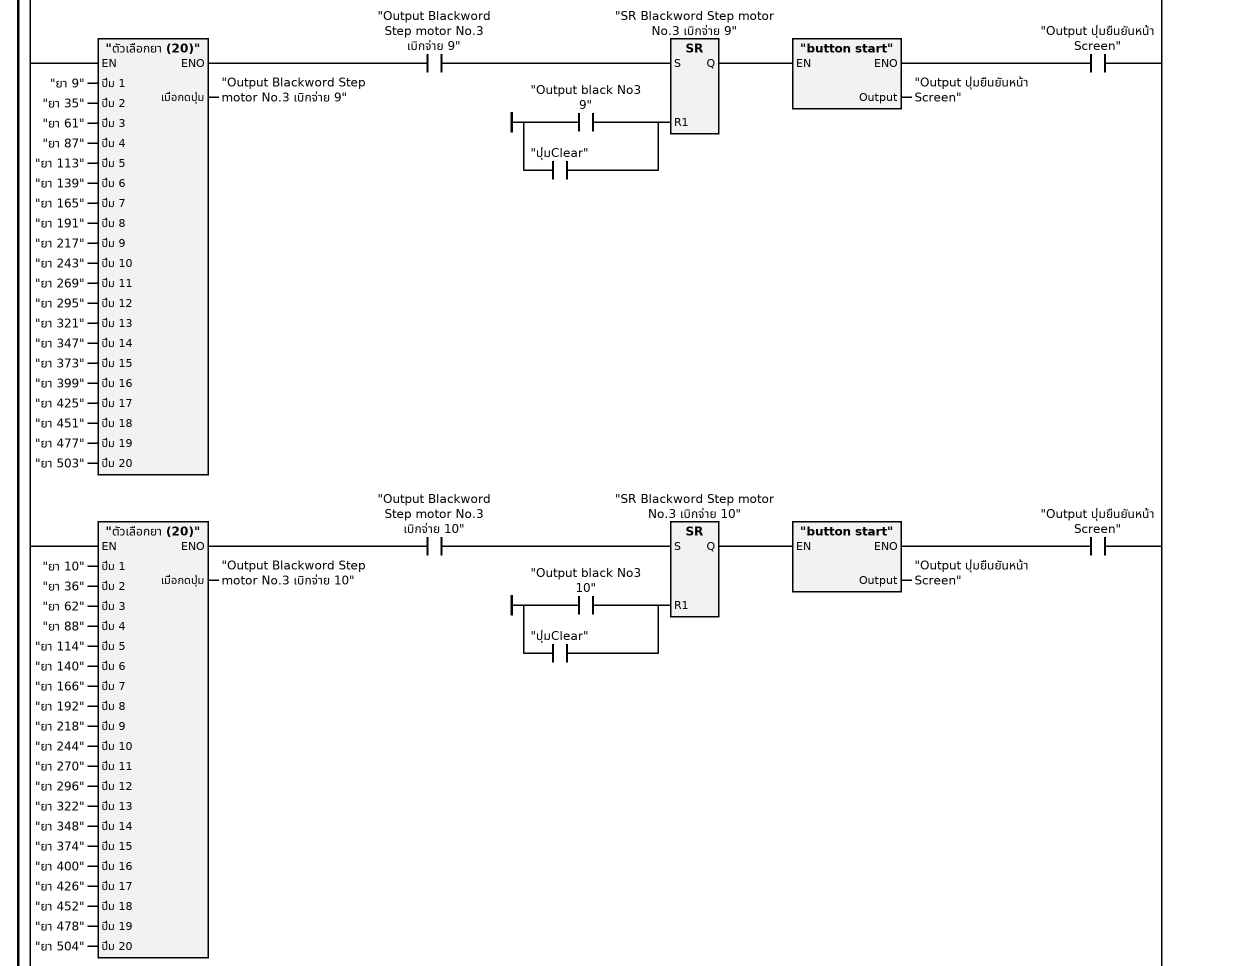
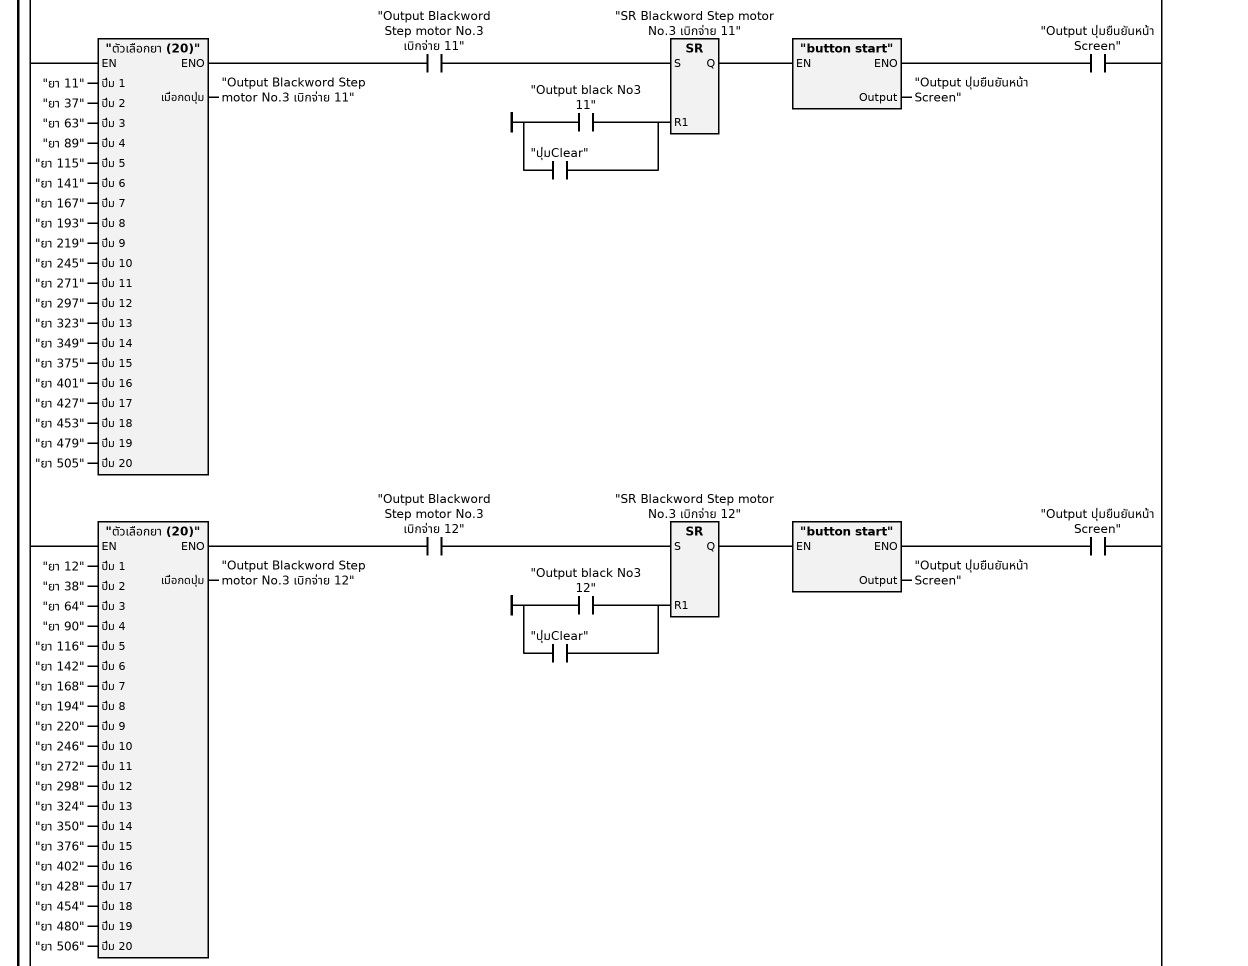
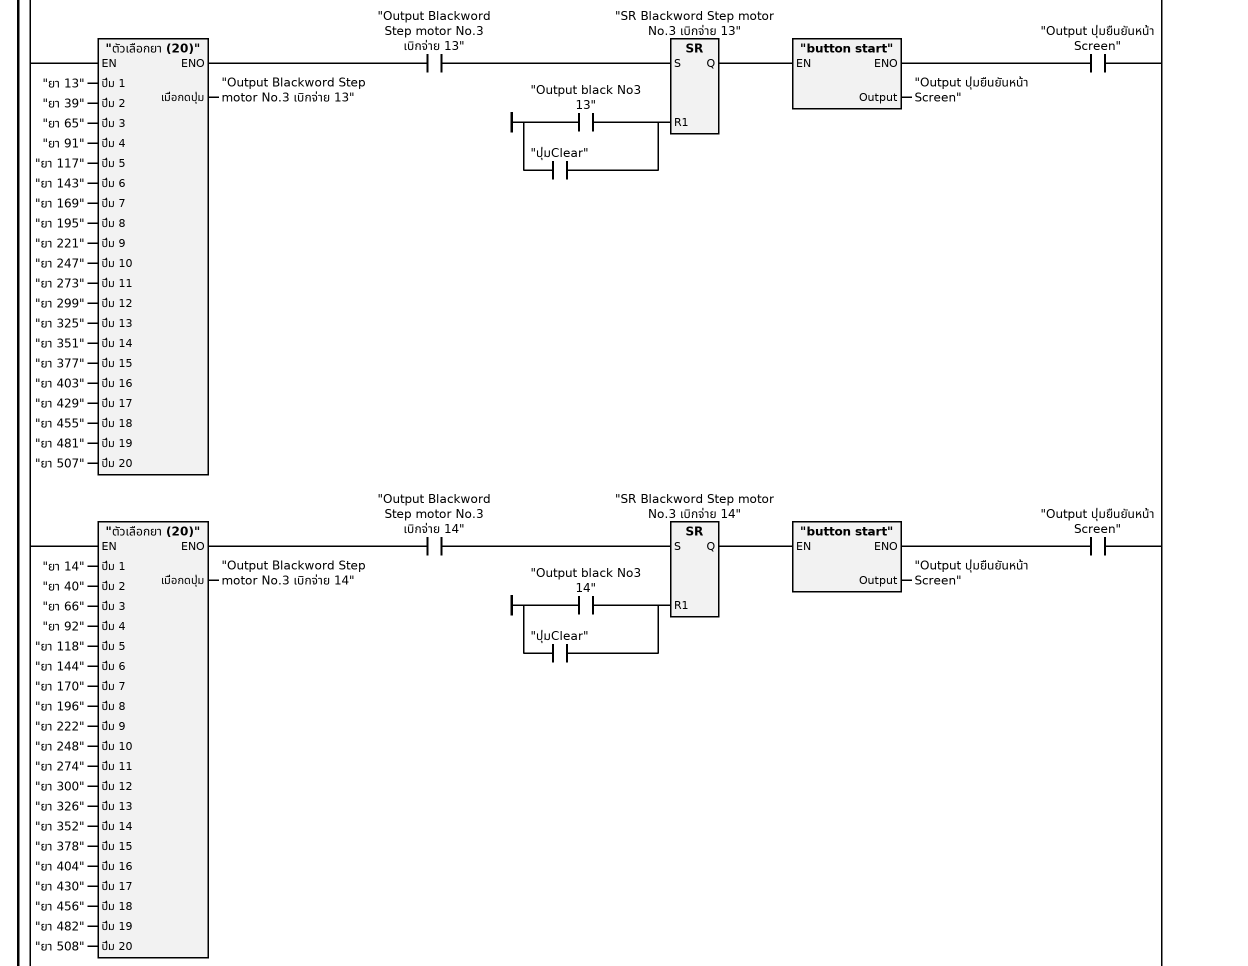
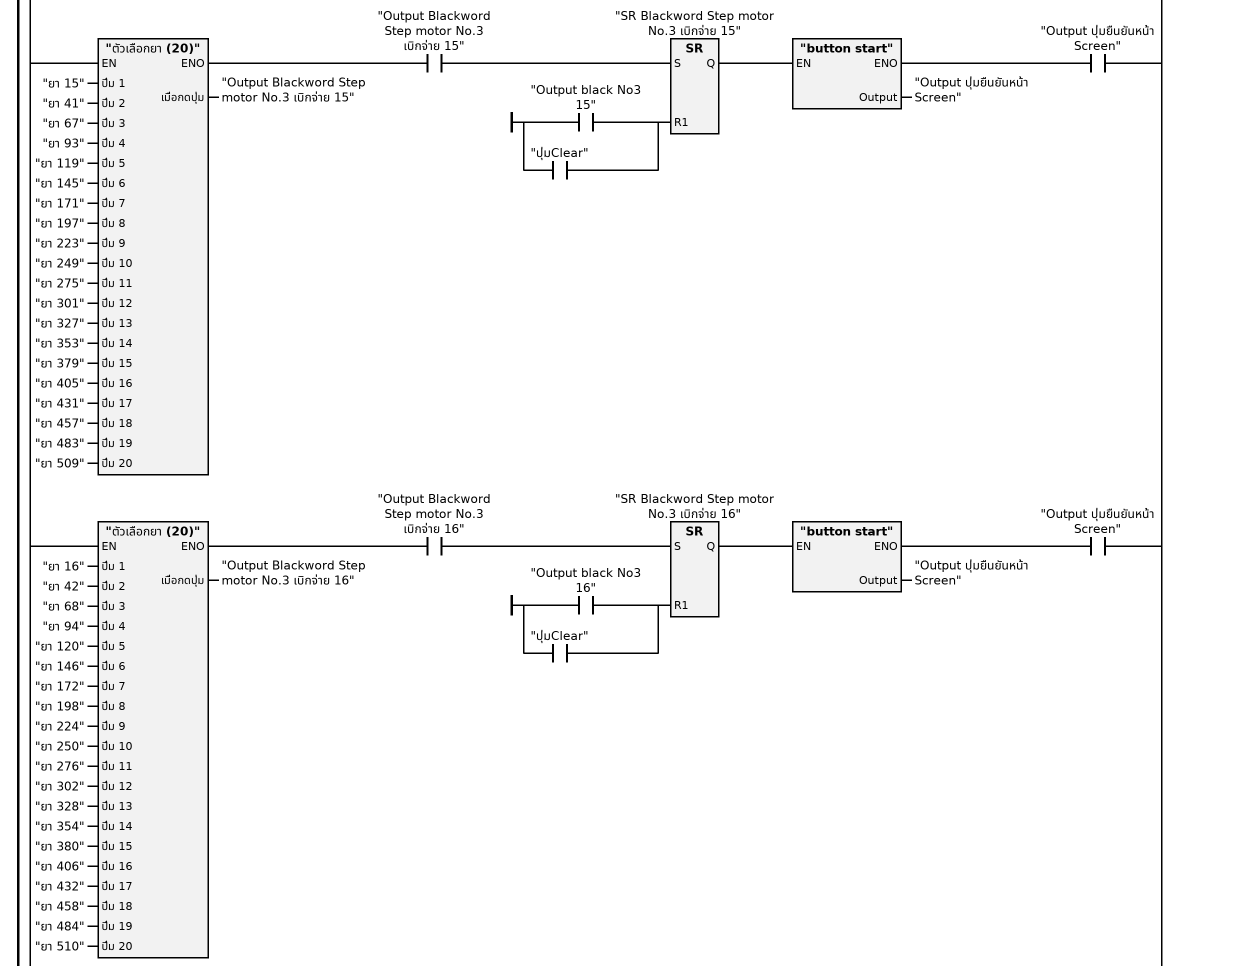
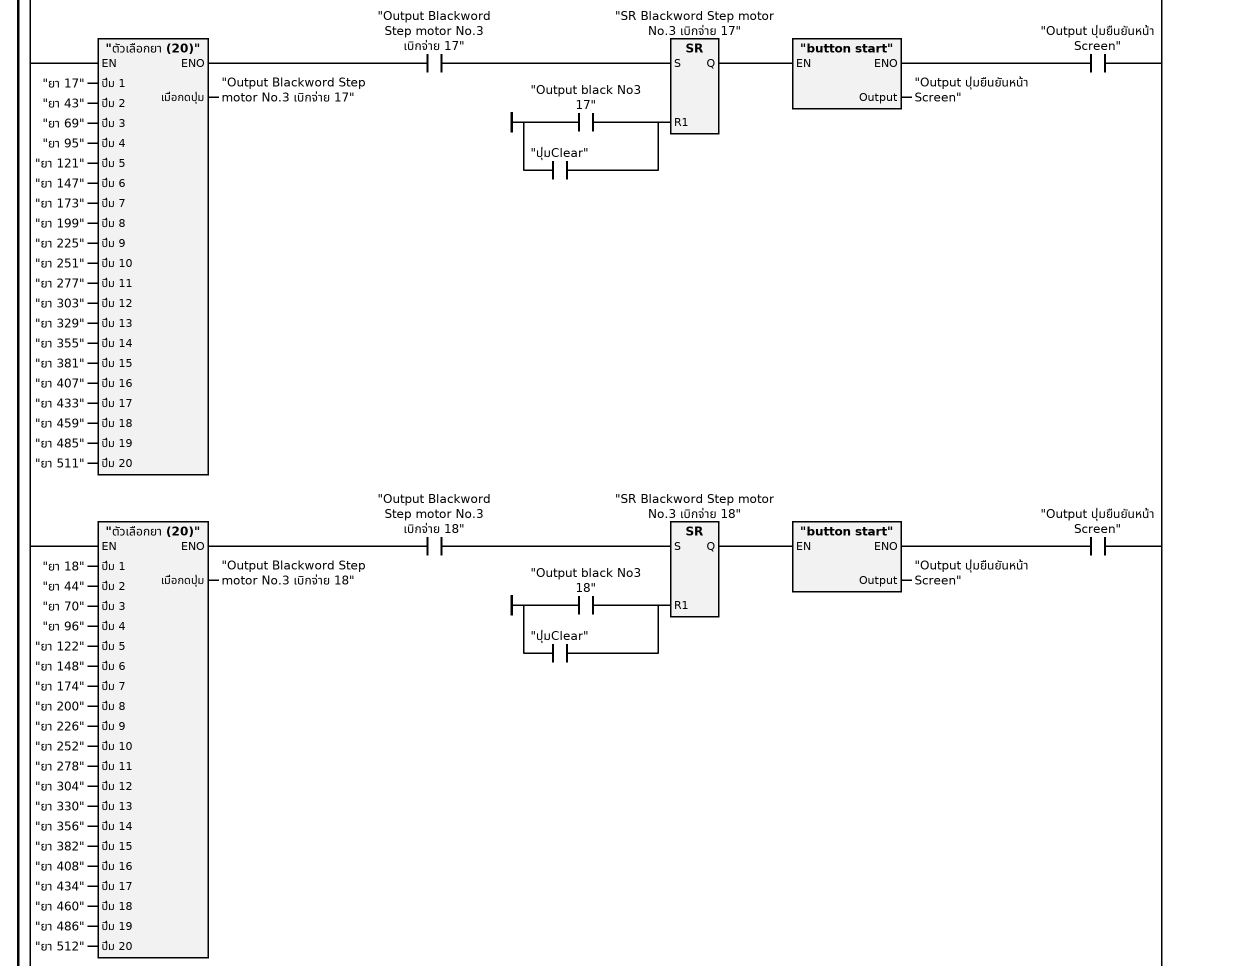
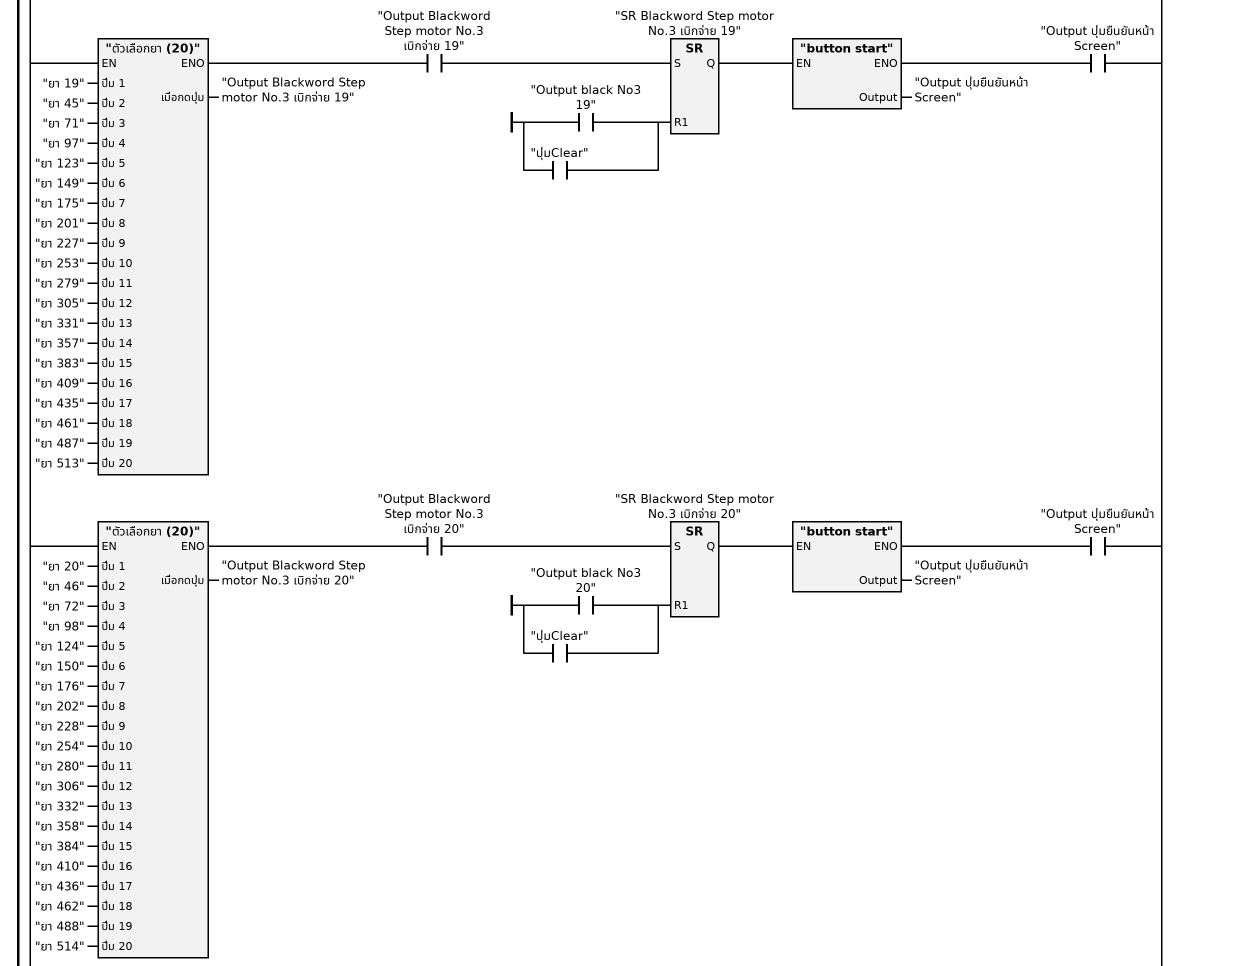
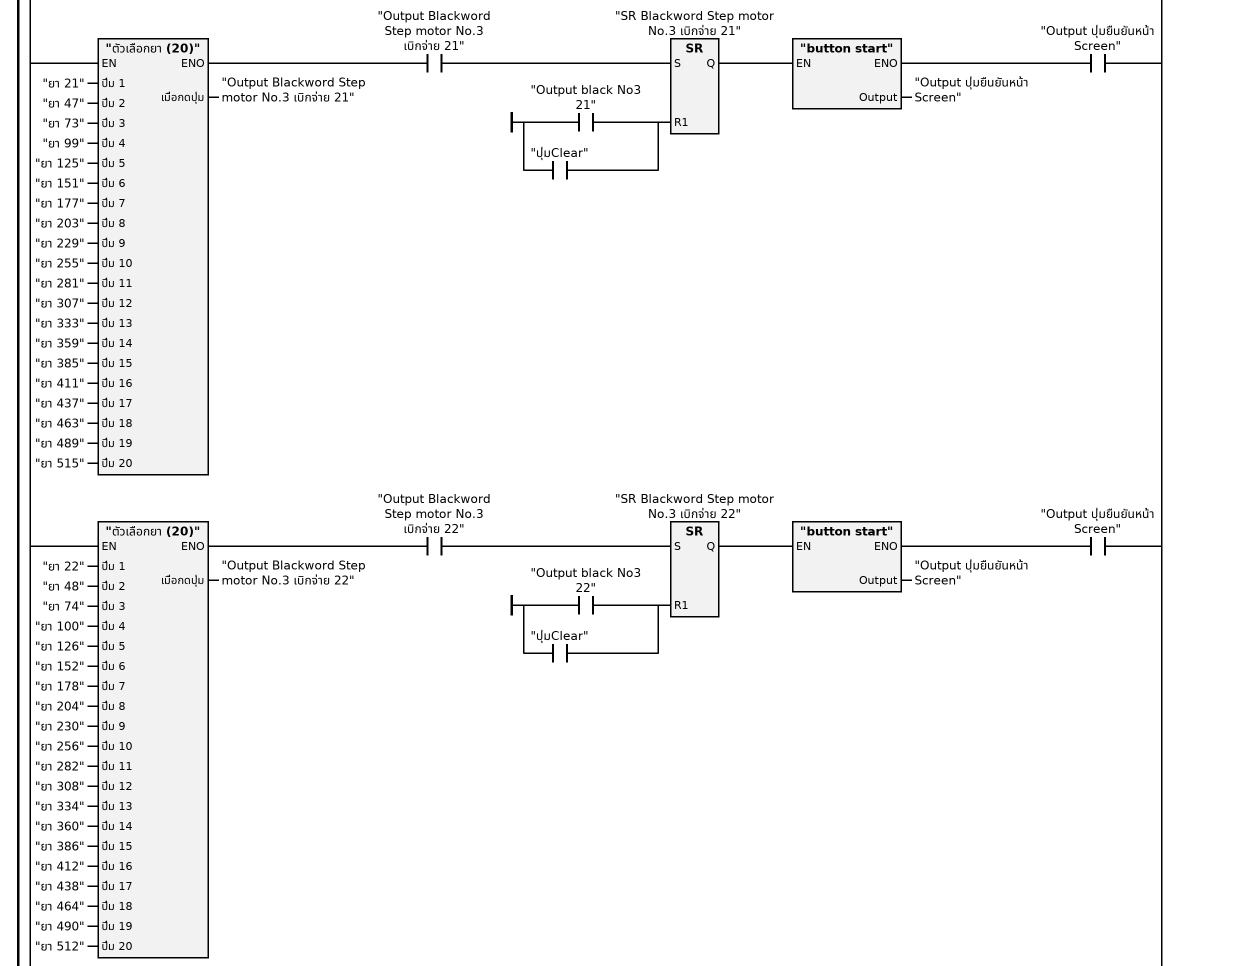
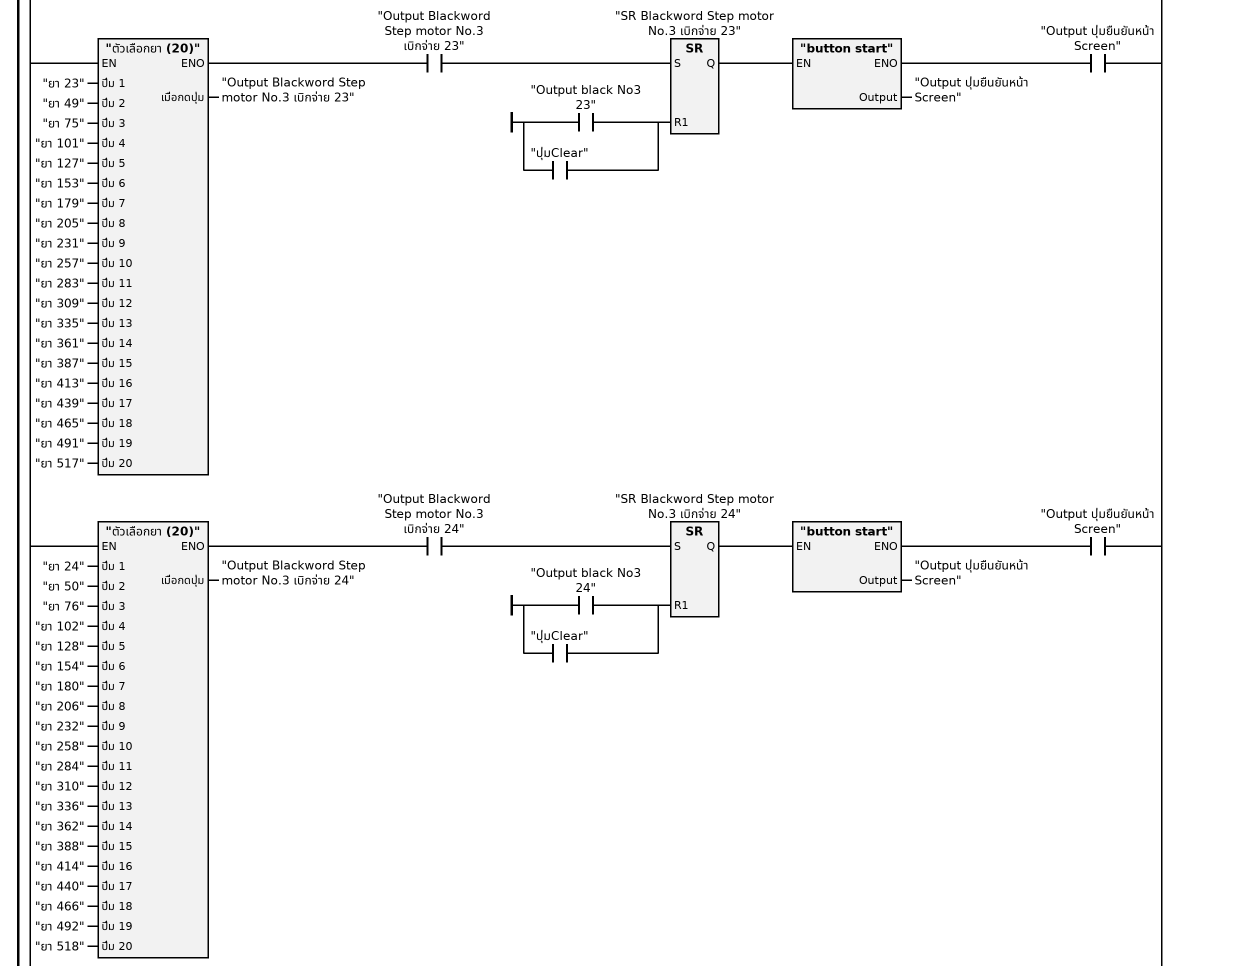
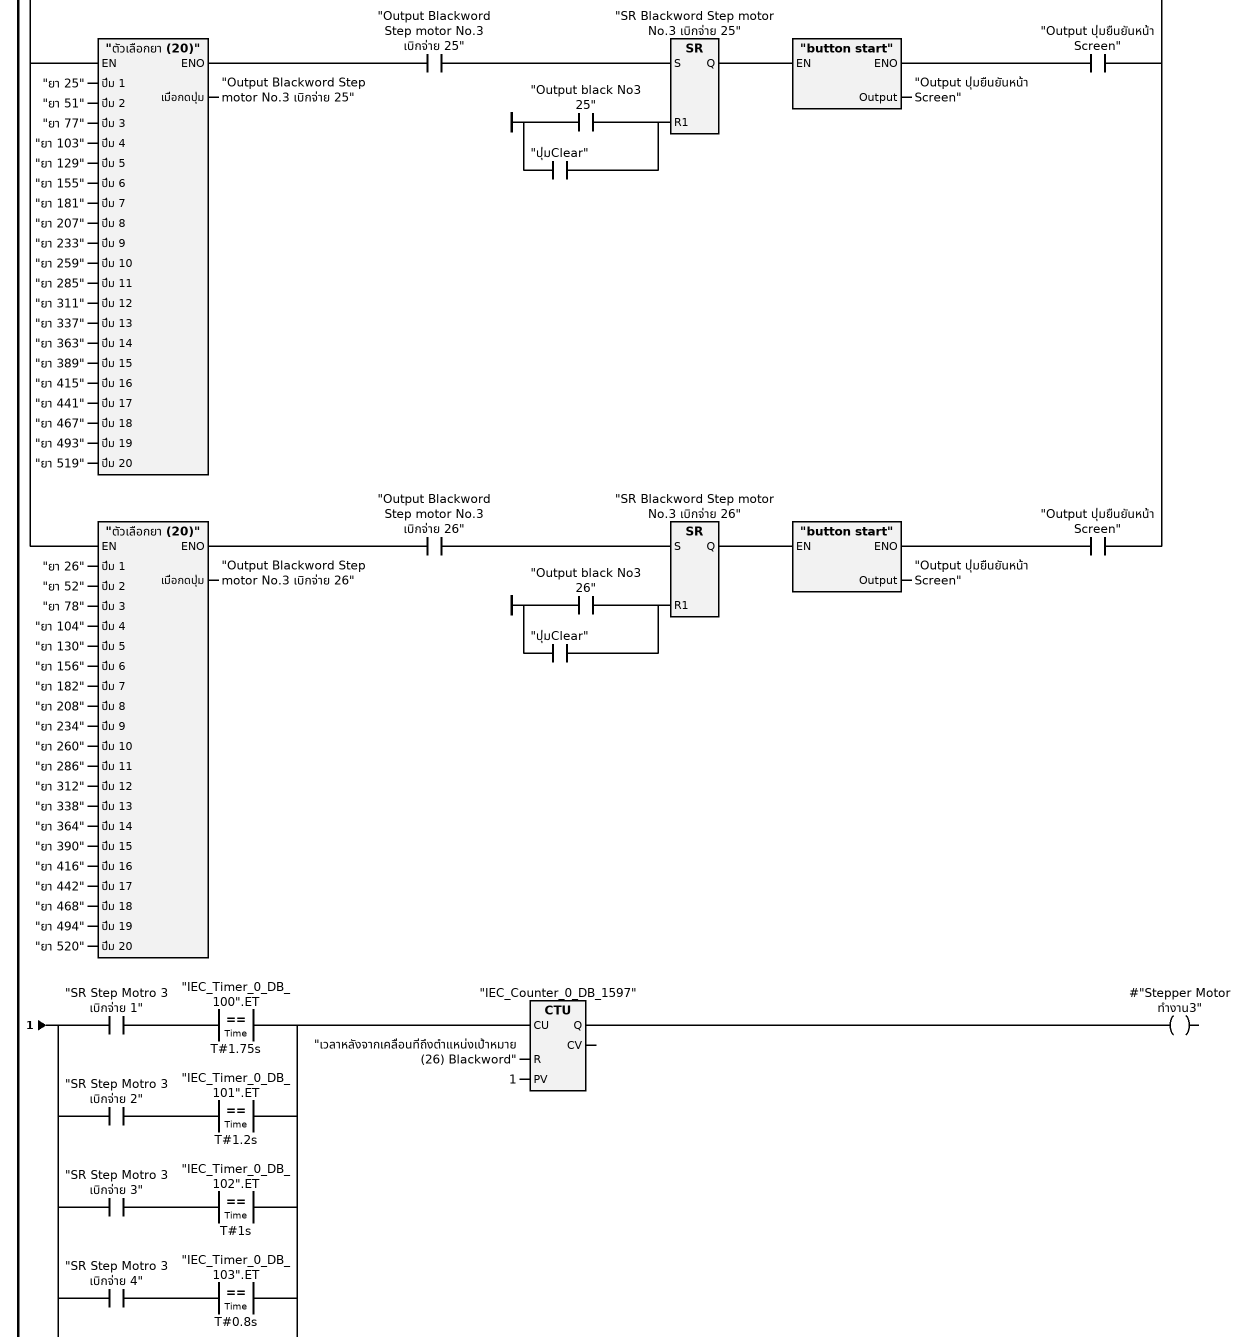
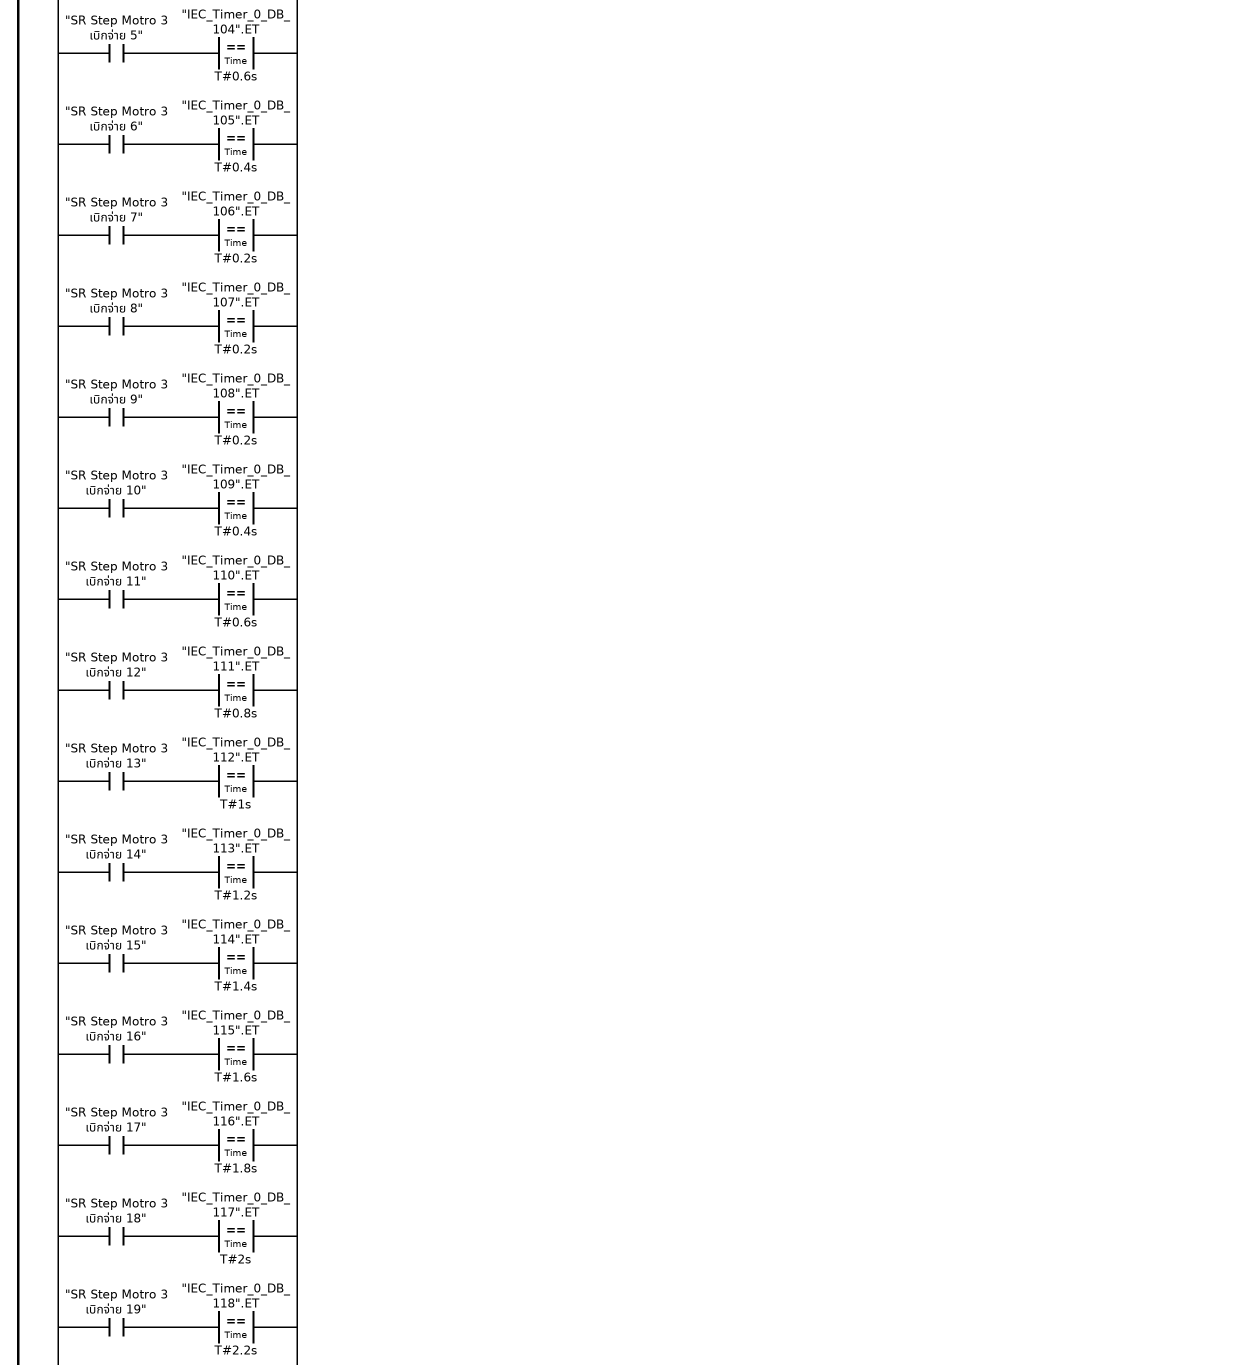
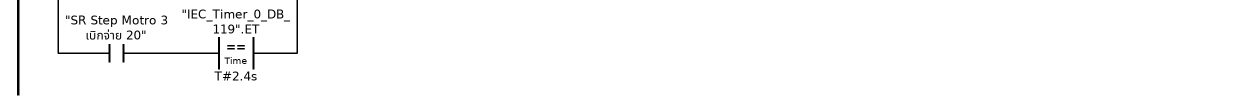
   "ตัวเลือกยา (20)"("ปึ่ม 1" := "ยา 1",
                     "ปึ่ม 2" := "ยา 27",
                     "ปึ่ม 3" := "ยา 53",
                     "ปึ่ม 4" := "ยา 79",
                     "ปึ่ม 5" := "ยา 105",
                     "ปึ่ม 6" := "ยา 131",
                     "ปึ่ม 7" := "ยา 157",
                     "ปึ่ม 8" := "ยา 183",
                     "ปึ่ม 9" := "ยา 209",
                     "ปึ่ม 10" := "ยา 235",
                     "ปึ่ม 11" := "ยา 261",
                     "ปึ่ม 12" := "ยา 287",
                     "ปึ่ม 13" := "ยา 313",
                     "ปึ่ม 14" := "ยา 339",
                     "ปึ่ม 15" := "ยา 365",
                     "ปึ่ม 16" := "ยา 391",
                     "ปึ่ม 17" := "ยา 417",
                     "ปึ่ม 18" := "ยา 443",
                     "ปึ่ม 19" := "ยา 469",
                     "ปึ่ม 20" := "ยา 495",
                     "เมื่อกดปุ่ม" => "Output Blackword Step motor No.3 เบิกจ่าย 1",
                     ENO => #_w1);
   IF #_w1 AND "Output Blackword Step motor No.3 เบิกจ่าย 1" THEN
       "SR Blackword Step motor No.3 เบิกจ่าย 1" := TRUE;   // SR flip-flop
   END_IF;
   IF "Output black No3 1" OR "ปุ่มClear" THEN "SR Blackword Step motor No.3 เบิกจ่าย 1" := FALSE; END_IF;
   "button start"(EN := "SR Blackword Step motor No.3 เบิกจ่าย 1",
                  Output => "Output ปุ่มยืนยันหน้า Screen",
                  ENO => #_w2);
   #_w4 := #_w2 AND "Output ปุ่มยืนยันหน้า Screen";
   "ตัวเลือกยา (20)"("ปึ่ม 1" := "ยา 2",
                     "ปึ่ม 2" := "ยา 28",
                     "ปึ่ม 3" := "ยา 54",
                     "ปึ่ม 4" := "ยา 80",
                     "ปึ่ม 5" := "ยา 106",
                     "ปึ่ม 6" := "ยา 132",
                     "ปึ่ม 7" := "ยา 158",
                     "ปึ่ม 8" := "ยา 184",
                     "ปึ่ม 9" := "ยา 201",
                     "ปึ่ม 10" := "ยา 236",
                     "ปึ่ม 11" := "ยา 262",
                     "ปึ่ม 12" := "ยา 288",
                     "ปึ่ม 13" := "ยา 314",
                     "ปึ่ม 14" := "ยา 340",
                     "ปึ่ม 15" := "ยา 366",
                     "ปึ่ม 16" := "ยา 392",
                     "ปึ่ม 17" := "ยา 418",
                     "ปึ่ม 18" := "ยา 444",
                     "ปึ่ม 19" := "ยา 470",
                     "ปึ่ม 20" := "ยา 492",
                     "เมื่อกดปุ่ม" => "Output Blackword Step motor No.3 เบิกจ่าย 2",
                     ENO => #_w3);
   IF #_w3 AND "Output Blackword Step motor No.3 เบิกจ่าย 2" THEN
       "SR Blackword Step motor No.3 เบิกจ่าย 2" := TRUE;   // SR flip-flop
   END_IF;
   IF "Output black No3 2" OR "ปุ่มClear" THEN "SR Blackword Step motor No.3 เบิกจ่าย 2" := FALSE; END_IF;
   "button start"(EN := "SR Blackword Step motor No.3 เบิกจ่าย 2",
                  Output => "Output ปุ่มยืนยันหน้า Screen",
                  ENO => #_w5);
   #_w7 := #_w5 AND "Output ปุ่มยืนยันหน้า Screen";
   "ตัวเลือกยา (20)"("ปึ่ม 1" := "ยา 3",
                     "ปึ่ม 2" := "ยา 29",
                     "ปึ่ม 3" := "ยา 55",
                     "ปึ่ม 4" := "ยา 81",
                     "ปึ่ม 5" := "ยา 107",
                     "ปึ่ม 6" := "ยา 133",
                     "ปึ่ม 7" := "ยา 159",
                     "ปึ่ม 8" := "ยา 185",
                     "ปึ่ม 9" := "ยา 211",
                     "ปึ่ม 10" := "ยา 237",
                     "ปึ่ม 11" := "ยา 263",
                     "ปึ่ม 12" := "ยา 289",
                     "ปึ่ม 13" := "ยา 315",
                     "ปึ่ม 14" := "ยา 341",
                     "ปึ่ม 15" := "ยา 367",
                     "ปึ่ม 16" := "ยา 393",
                     "ปึ่ม 17" := "ยา 419",
                     "ปึ่ม 18" := "ยา 445",
                     "ปึ่ม 19" := "ยา 471",
                     "ปึ่ม 20" := "ยา 497",
                     "เมื่อกดปุ่ม" => "Output Blackword Step motor No.3 เบิกจ่าย 3",
                     ENO => #_w6);
   IF #_w6 AND "Output Blackword Step motor No.3 เบิกจ่าย 3" THEN
       "SR Blackword Step motor No.3 เบิกจ่าย 3" := TRUE;   // SR flip-flop
   END_IF;
   IF "Output black No3 3" OR "ปุ่มClear" THEN "SR Blackword Step motor No.3 เบิกจ่าย 3" := FALSE; END_IF;
   "button start"(EN := "SR Blackword Step motor No.3 เบิกจ่าย 3",
                  Output => "Output ปุ่มยืนยันหน้า Screen",
                  ENO => #_w8);
   #_w10 := #_w8 AND "Output ปุ่มยืนยันหน้า Screen";
   "ตัวเลือกยา (20)"("ปึ่ม 1" := "ยา 4",
                     "ปึ่ม 2" := "ยา 30",
                     "ปึ่ม 3" := "ยา 56",
                     "ปึ่ม 4" := "ยา 82",
                     "ปึ่ม 5" := "ยา 108",
                     "ปึ่ม 6" := "ยา 134",
                     "ปึ่ม 7" := "ยา 160",
                     "ปึ่ม 8" := "ยา 186",
                     "ปึ่ม 9" := "ยา 212",
                     "ปึ่ม 10" := "ยา 238",
                     "ปึ่ม 11" := "ยา 264",
                     "ปึ่ม 12" := "ยา 290",
                     "ปึ่ม 13" := "ยา 316",
                     "ปึ่ม 14" := "ยา 342",
                     "ปึ่ม 15" := "ยา 368",
                     "ปึ่ม 16" := "ยา 394",
                     "ปึ่ม 17" := "ยา 420",
                     "ปึ่ม 18" := "ยา 446",
                     "ปึ่ม 19" := "ยา 472",
                     "ปึ่ม 20" := "ยา 498",
                     "เมื่อกดปุ่ม" => "Output Blackword Step motor No.3 เบิกจ่าย 4",
                     ENO => #_w9);
   IF #_w9 AND "Output Blackword Step motor No.3 เบิกจ่าย 4" THEN
       "SR Blackword Step motor No.3 เบิกจ่าย 4" := TRUE;   // SR flip-flop
   END_IF;
   IF "Output black No3 4" OR "ปุ่มClear" THEN "SR Blackword Step motor No.3 เบิกจ่าย 4" := FALSE; END_IF;
   "button start"(EN := "SR Blackword Step motor No.3 เบิกจ่าย 4",
                  Output => "Output ปุ่มยืนยันหน้า Screen",
                  ENO => #_w11);
   #_w13 := #_w11 AND "Output ปุ่มยืนยันหน้า Screen";
   "ตัวเลือกยา (20)"("ปึ่ม 1" := "ยา 5",
                     "ปึ่ม 2" := "ยา 31",
                     "ปึ่ม 3" := "ยา 57",
                     "ปึ่ม 4" := "ยา 83",
                     "ปึ่ม 5" := "ยา 109",
                     "ปึ่ม 6" := "ยา 135",
                     "ปึ่ม 7" := "ยา 161",
                     "ปึ่ม 8" := "ยา 187",
                     "ปึ่ม 9" := "ยา 213",
                     "ปึ่ม 10" := "ยา 239",
                     "ปึ่ม 11" := "ยา 265",
                     "ปึ่ม 12" := "ยา 291",
                     "ปึ่ม 13" := "ยา 317",
                     "ปึ่ม 14" := "ยา 343",
                     "ปึ่ม 15" := "ยา 369",
                     "ปึ่ม 16" := "ยา 395",
                     "ปึ่ม 17" := "ยา 421",
                     "ปึ่ม 18" := "ยา 447",
                     "ปึ่ม 19" := "ยา 473",
                     "ปึ่ม 20" := "ยา 499",
                     "เมื่อกดปุ่ม" => "Output Blackword Step motor No.3 เบิกจ่าย 5",
                     ENO => #_w12);
   IF #_w12 AND "Output Blackword Step motor No.3 เบิกจ่าย 5" THEN
       "SR Blackword Step motor No.3 เบิกจ่าย 5" := TRUE;   // SR flip-flop
   END_IF;
   IF "Output black No3 5" OR "ปุ่มClear" THEN "SR Blackword Step motor No.3 เบิกจ่าย 5" := FALSE; END_IF;
   "button start"(EN := "SR Blackword Step motor No.3 เบิกจ่าย 5",
                  Output => "Output ปุ่มยืนยันหน้า Screen",
                  ENO => #_w14);
   #_w16 := #_w14 AND "Output ปุ่มยืนยันหน้า Screen";
   "ตัวเลือกยา (20)"("ปึ่ม 1" := "ยา 6",
                     "ปึ่ม 2" := "ยา 32",
                     "ปึ่ม 3" := "ยา 58",
                     "ปึ่ม 4" := "ยา 84",
                     "ปึ่ม 5" := "ยา 110",
                     "ปึ่ม 6" := "ยา 136",
                     "ปึ่ม 7" := "ยา 162",
                     "ปึ่ม 8" := "ยา 188",
                     "ปึ่ม 9" := "ยา 214",
                     "ปึ่ม 10" := "ยา 240",
                     "ปึ่ม 11" := "ยา 266",
                     "ปึ่ม 12" := "ยา 292",
                     "ปึ่ม 13" := "ยา 318",
                     "ปึ่ม 14" := "ยา 344",
                     "ปึ่ม 15" := "ยา 370",
                     "ปึ่ม 16" := "ยา 396",
                     "ปึ่ม 17" := "ยา 422",
                     "ปึ่ม 18" := "ยา 448",
                     "ปึ่ม 19" := "ยา 474",
                     "ปึ่ม 20" := "ยา 500",
                     "เมื่อกดปุ่ม" => "Output Blackword Step motor No.3 เบิกจ่าย 6",
                     ENO => #_w15);
   IF #_w15 AND "Output Blackword Step motor No.3 เบิกจ่าย 6" THEN
       "SR Blackword Step motor No.3 เบิกจ่าย 6" := TRUE;   // SR flip-flop
   END_IF;
   IF "Output black No3 6" OR "ปุ่มClear" THEN "SR Blackword Step motor No.3 เบิกจ่าย 6" := FALSE; END_IF;
   "button start"(EN := "SR Blackword Step motor No.3 เบิกจ่าย 6",
                  Output => "Output ปุ่มยืนยันหน้า Screen",
                  ENO => #_w17);
   #_w19 := #_w17 AND "Output ปุ่มยืนยันหน้า Screen";
   "ตัวเลือกยา (20)"("ปึ่ม 1" := "ยา 7",
                     "ปึ่ม 2" := "ยา 33",
                     "ปึ่ม 3" := "ยา 59",
                     "ปึ่ม 4" := "ยา 85",
                     "ปึ่ม 5" := "ยา 111",
                     "ปึ่ม 6" := "ยา 137",
                     "ปึ่ม 7" := "ยา 163",
                     "ปึ่ม 8" := "ยา 189",
                     "ปึ่ม 9" := "ยา 215",
                     "ปึ่ม 10" := "ยา 241",
                     "ปึ่ม 11" := "ยา 267",
                     "ปึ่ม 12" := "ยา 293",
                     "ปึ่ม 13" := "ยา 319",
                     "ปึ่ม 14" := "ยา 345",
                     "ปึ่ม 15" := "ยา 371",
                     "ปึ่ม 16" := "ยา 397",
                     "ปึ่ม 17" := "ยา 423",
                     "ปึ่ม 18" := "ยา 449",
                     "ปึ่ม 19" := "ยา 475",
                     "ปึ่ม 20" := "ยา 501",
                     "เมื่อกดปุ่ม" => "Output Blackword Step motor No.3 เบิกจ่าย 7",
                     ENO => #_w18);
   IF #_w18 AND "Output Blackword Step motor No.3 เบิกจ่าย 7" THEN
       "SR Blackword Step motor No.3 เบิกจ่าย 7" := TRUE;   // SR flip-flop
   END_IF;
   IF "Output black No3 7" OR "ปุ่มClear" THEN "SR Blackword Step motor No.3 เบิกจ่าย 7" := FALSE; END_IF;
   "button start"(EN := "SR Blackword Step motor No.3 เบิกจ่าย 7",
                  Output => "Output ปุ่มยืนยันหน้า Screen",
                  ENO => #_w20);
   #_w22 := #_w20 AND "Output ปุ่มยืนยันหน้า Screen";
   "ตัวเลือกยา (20)"("ปึ่ม 1" := "ยา 8",
                     "ปึ่ม 2" := "ยา 34",
                     "ปึ่ม 3" := "ยา 60",
                     "ปึ่ม 4" := "ยา 86",
                     "ปึ่ม 5" := "ยา 112",
                     "ปึ่ม 6" := "ยา 138",
                     "ปึ่ม 7" := "ยา 164",
                     "ปึ่ม 8" := "ยา 190",
                     "ปึ่ม 9" := "ยา 216",
                     "ปึ่ม 10" := "ยา 242",
                     "ปึ่ม 11" := "ยา 268",
                     "ปึ่ม 12" := "ยา 294",
                     "ปึ่ม 13" := "ยา 320",
                     "ปึ่ม 14" := "ยา 346",
                     "ปึ่ม 15" := "ยา 372",
                     "ปึ่ม 16" := "ยา 398",
                     "ปึ่ม 17" := "ยา 424",
                     "ปึ่ม 18" := "ยา 450",
                     "ปึ่ม 19" := "ยา 476",
                     "ปึ่ม 20" := "ยา 502",
                     "เมื่อกดปุ่ม" => "Output Blackword Step motor No.3 เบิกจ่าย 8",
                     ENO => #_w21);
   IF #_w21 AND "Output Blackword Step motor No.3 เบิกจ่าย 8" THEN
       "SR Blackword Step motor No.3 เบิกจ่าย 8" := TRUE;   // SR flip-flop
   END_IF;
   IF "Output black No3 8" OR "ปุ่มClear" THEN "SR Blackword Step motor No.3 เบิกจ่าย 8" := FALSE; END_IF;
   "button start"(EN := "SR Blackword Step motor No.3 เบิกจ่าย 8",
                  Output => "Output ปุ่มยืนยันหน้า Screen",
                  ENO => #_w23);
   #_w25 := #_w23 AND "Output ปุ่มยืนยันหน้า Screen";
   "ตัวเลือกยา (20)"("ปึ่ม 1" := "ยา 9",
                     "ปึ่ม 2" := "ยา 35",
                     "ปึ่ม 3" := "ยา 61",
                     "ปึ่ม 4" := "ยา 87",
                     "ปึ่ม 5" := "ยา 113",
                     "ปึ่ม 6" := "ยา 139",
                     "ปึ่ม 7" := "ยา 165",
                     "ปึ่ม 8" := "ยา 191",
                     "ปึ่ม 9" := "ยา 217",
                     "ปึ่ม 10" := "ยา 243",
                     "ปึ่ม 11" := "ยา 269",
                     "ปึ่ม 12" := "ยา 295",
                     "ปึ่ม 13" := "ยา 321",
                     "ปึ่ม 14" := "ยา 347",
                     "ปึ่ม 15" := "ยา 373",
                     "ปึ่ม 16" := "ยา 399",
                     "ปึ่ม 17" := "ยา 425",
                     "ปึ่ม 18" := "ยา 451",
                     "ปึ่ม 19" := "ยา 477",
                     "ปึ่ม 20" := "ยา 503",
                     "เมื่อกดปุ่ม" => "Output Blackword Step motor No.3 เบิกจ่าย 9",
                     ENO => #_w24);
   IF #_w24 AND "Output Blackword Step motor No.3 เบิกจ่าย 9" THEN
       "SR Blackword Step motor No.3 เบิกจ่าย 9" := TRUE;   // SR flip-flop
   END_IF;
   IF "Output black No3 9" OR "ปุ่มClear" THEN "SR Blackword Step motor No.3 เบิกจ่าย 9" := FALSE; END_IF;
   "button start"(EN := "SR Blackword Step motor No.3 เบิกจ่าย 9",
                  Output => "Output ปุ่มยืนยันหน้า Screen",
                  ENO => #_w26);
   #_w28 := #_w26 AND "Output ปุ่มยืนยันหน้า Screen";
   "ตัวเลือกยา (20)"("ปึ่ม 1" := "ยา 10",
                     "ปึ่ม 2" := "ยา 36",
                     "ปึ่ม 3" := "ยา 62",
                     "ปึ่ม 4" := "ยา 88",
                     "ปึ่ม 5" := "ยา 114",
                     "ปึ่ม 6" := "ยา 140",
                     "ปึ่ม 7" := "ยา 166",
                     "ปึ่ม 8" := "ยา 192",
                     "ปึ่ม 9" := "ยา 218",
                     "ปึ่ม 10" := "ยา 244",
                     "ปึ่ม 11" := "ยา 270",
                     "ปึ่ม 12" := "ยา 296",
                     "ปึ่ม 13" := "ยา 322",
                     "ปึ่ม 14" := "ยา 348",
                     "ปึ่ม 15" := "ยา 374",
                     "ปึ่ม 16" := "ยา 400",
                     "ปึ่ม 17" := "ยา 426",
                     "ปึ่ม 18" := "ยา 452",
                     "ปึ่ม 19" := "ยา 478",
                     "ปึ่ม 20" := "ยา 504",
                     "เมื่อกดปุ่ม" => "Output Blackword Step motor No.3 เบิกจ่าย 10",
                     ENO => #_w27);
   IF #_w27 AND "Output Blackword Step motor No.3 เบิกจ่าย 10" THEN
       "SR Blackword Step motor No.3 เบิกจ่าย 10" := TRUE;   // SR flip-flop
   END_IF;
   IF "Output black No3 10" OR "ปุ่มClear" THEN "SR Blackword Step motor No.3 เบิกจ่าย 10" := FALSE; END_IF;
   "button start"(EN := "SR Blackword Step motor No.3 เบิกจ่าย 10",
                  Output => "Output ปุ่มยืนยันหน้า Screen",
                  ENO => #_w29);
   #_w31 := #_w29 AND "Output ปุ่มยืนยันหน้า Screen";
   "ตัวเลือกยา (20)"("ปึ่ม 1" := "ยา 11",
                     "ปึ่ม 2" := "ยา 37",
                     "ปึ่ม 3" := "ยา 63",
                     "ปึ่ม 4" := "ยา 89",
                     "ปึ่ม 5" := "ยา 115",
                     "ปึ่ม 6" := "ยา 141",
                     "ปึ่ม 7" := "ยา 167",
                     "ปึ่ม 8" := "ยา 193",
                     "ปึ่ม 9" := "ยา 219",
                     "ปึ่ม 10" := "ยา 245",
                     "ปึ่ม 11" := "ยา 271",
                     "ปึ่ม 12" := "ยา 297",
                     "ปึ่ม 13" := "ยา 323",
                     "ปึ่ม 14" := "ยา 349",
                     "ปึ่ม 15" := "ยา 375",
                     "ปึ่ม 16" := "ยา 401",
                     "ปึ่ม 17" := "ยา 427",
                     "ปึ่ม 18" := "ยา 453",
                     "ปึ่ม 19" := "ยา 479",
                     "ปึ่ม 20" := "ยา 505",
                     "เมื่อกดปุ่ม" => "Output Blackword Step motor No.3 เบิกจ่าย 11",
                     ENO => #_w30);
   IF #_w30 AND "Output Blackword Step motor No.3 เบิกจ่าย 11" THEN
       "SR Blackword Step motor No.3 เบิกจ่าย 11" := TRUE;   // SR flip-flop
   END_IF;
   IF "Output black No3 11" OR "ปุ่มClear" THEN "SR Blackword Step motor No.3 เบิกจ่าย 11" := FALSE; END_IF;
   "button start"(EN := "SR Blackword Step motor No.3 เบิกจ่าย 11",
                  Output => "Output ปุ่มยืนยันหน้า Screen",
                  ENO => #_w32);
   #_w34 := #_w32 AND "Output ปุ่มยืนยันหน้า Screen";
   "ตัวเลือกยา (20)"("ปึ่ม 1" := "ยา 12",
                     "ปึ่ม 2" := "ยา 38",
                     "ปึ่ม 3" := "ยา 64",
                     "ปึ่ม 4" := "ยา 90",
                     "ปึ่ม 5" := "ยา 116",
                     "ปึ่ม 6" := "ยา 142",
                     "ปึ่ม 7" := "ยา 168",
                     "ปึ่ม 8" := "ยา 194",
                     "ปึ่ม 9" := "ยา 220",
                     "ปึ่ม 10" := "ยา 246",
                     "ปึ่ม 11" := "ยา 272",
                     "ปึ่ม 12" := "ยา 298",
                     "ปึ่ม 13" := "ยา 324",
                     "ปึ่ม 14" := "ยา 350",
                     "ปึ่ม 15" := "ยา 376",
                     "ปึ่ม 16" := "ยา 402",
                     "ปึ่ม 17" := "ยา 428",
                     "ปึ่ม 18" := "ยา 454",
                     "ปึ่ม 19" := "ยา 480",
                     "ปึ่ม 20" := "ยา 506",
                     "เมื่อกดปุ่ม" => "Output Blackword Step motor No.3 เบิกจ่าย 12",
                     ENO => #_w33);
   IF #_w33 AND "Output Blackword Step motor No.3 เบิกจ่าย 12" THEN
       "SR Blackword Step motor No.3 เบิกจ่าย 12" := TRUE;   // SR flip-flop
   END_IF;
   IF "Output black No3 12" OR "ปุ่มClear" THEN "SR Blackword Step motor No.3 เบิกจ่าย 12" := FALSE; END_IF;
   "button start"(EN := "SR Blackword Step motor No.3 เบิกจ่าย 12",
                  Output => "Output ปุ่มยืนยันหน้า Screen",
                  ENO => #_w35);
   #_w37 := #_w35 AND "Output ปุ่มยืนยันหน้า Screen";
   "ตัวเลือกยา (20)"("ปึ่ม 1" := "ยา 13",
                     "ปึ่ม 2" := "ยา 39",
                     "ปึ่ม 3" := "ยา 65",
                     "ปึ่ม 4" := "ยา 91",
                     "ปึ่ม 5" := "ยา 117",
                     "ปึ่ม 6" := "ยา 143",
                     "ปึ่ม 7" := "ยา 169",
                     "ปึ่ม 8" := "ยา 195",
                     "ปึ่ม 9" := "ยา 221",
                     "ปึ่ม 10" := "ยา 247",
                     "ปึ่ม 11" := "ยา 273",
                     "ปึ่ม 12" := "ยา 299",
                     "ปึ่ม 13" := "ยา 325",
                     "ปึ่ม 14" := "ยา 351",
                     "ปึ่ม 15" := "ยา 377",
                     "ปึ่ม 16" := "ยา 403",
                     "ปึ่ม 17" := "ยา 429",
                     "ปึ่ม 18" := "ยา 455",
                     "ปึ่ม 19" := "ยา 481",
                     "ปึ่ม 20" := "ยา 507",
                     "เมื่อกดปุ่ม" => "Output Blackword Step motor No.3 เบิกจ่าย 13",
                     ENO => #_w36);
   IF #_w36 AND "Output Blackword Step motor No.3 เบิกจ่าย 13" THEN
       "SR Blackword Step motor No.3 เบิกจ่าย 13" := TRUE;   // SR flip-flop
   END_IF;
   IF "Output black No3 13" OR "ปุ่มClear" THEN "SR Blackword Step motor No.3 เบิกจ่าย 13" := FALSE; END_IF;
   "button start"(EN := "SR Blackword Step motor No.3 เบิกจ่าย 13",
                  Output => "Output ปุ่มยืนยันหน้า Screen",
                  ENO => #_w38);
   #_w40 := #_w38 AND "Output ปุ่มยืนยันหน้า Screen";
   "ตัวเลือกยา (20)"("ปึ่ม 1" := "ยา 14",
                     "ปึ่ม 2" := "ยา 40",
                     "ปึ่ม 3" := "ยา 66",
                     "ปึ่ม 4" := "ยา 92",
                     "ปึ่ม 5" := "ยา 118",
                     "ปึ่ม 6" := "ยา 144",
                     "ปึ่ม 7" := "ยา 170",
                     "ปึ่ม 8" := "ยา 196",
                     "ปึ่ม 9" := "ยา 222",
                     "ปึ่ม 10" := "ยา 248",
                     "ปึ่ม 11" := "ยา 274",
                     "ปึ่ม 12" := "ยา 300",
                     "ปึ่ม 13" := "ยา 326",
                     "ปึ่ม 14" := "ยา 352",
                     "ปึ่ม 15" := "ยา 378",
                     "ปึ่ม 16" := "ยา 404",
                     "ปึ่ม 17" := "ยา 430",
                     "ปึ่ม 18" := "ยา 456",
                     "ปึ่ม 19" := "ยา 482",
                     "ปึ่ม 20" := "ยา 508",
                     "เมื่อกดปุ่ม" => "Output Blackword Step motor No.3 เบิกจ่าย 14",
                     ENO => #_w39);
   IF #_w39 AND "Output Blackword Step motor No.3 เบิกจ่าย 14" THEN
       "SR Blackword Step motor No.3 เบิกจ่าย 14" := TRUE;   // SR flip-flop
   END_IF;
   IF "Output black No3 14" OR "ปุ่มClear" THEN "SR Blackword Step motor No.3 เบิกจ่าย 14" := FALSE; END_IF;
   "button start"(EN := "SR Blackword Step motor No.3 เบิกจ่าย 14",
                  Output => "Output ปุ่มยืนยันหน้า Screen",
                  ENO => #_w41);
   #_w43 := #_w41 AND "Output ปุ่มยืนยันหน้า Screen";
   "ตัวเลือกยา (20)"("ปึ่ม 1" := "ยา 15",
                     "ปึ่ม 2" := "ยา 41",
                     "ปึ่ม 3" := "ยา 67",
                     "ปึ่ม 4" := "ยา 93",
                     "ปึ่ม 5" := "ยา 119",
                     "ปึ่ม 6" := "ยา 145",
                     "ปึ่ม 7" := "ยา 171",
                     "ปึ่ม 8" := "ยา 197",
                     "ปึ่ม 9" := "ยา 223",
                     "ปึ่ม 10" := "ยา 249",
                     "ปึ่ม 11" := "ยา 275",
                     "ปึ่ม 12" := "ยา 301",
                     "ปึ่ม 13" := "ยา 327",
                     "ปึ่ม 14" := "ยา 353",
                     "ปึ่ม 15" := "ยา 379",
                     "ปึ่ม 16" := "ยา 405",
                     "ปึ่ม 17" := "ยา 431",
                     "ปึ่ม 18" := "ยา 457",
                     "ปึ่ม 19" := "ยา 483",
                     "ปึ่ม 20" := "ยา 509",
                     "เมื่อกดปุ่ม" => "Output Blackword Step motor No.3 เบิกจ่าย 15",
                     ENO => #_w42);
   IF #_w42 AND "Output Blackword Step motor No.3 เบิกจ่าย 15" THEN
       "SR Blackword Step motor No.3 เบิกจ่าย 15" := TRUE;   // SR flip-flop
   END_IF;
   IF "Output black No3 15" OR "ปุ่มClear" THEN "SR Blackword Step motor No.3 เบิกจ่าย 15" := FALSE; END_IF;
   "button start"(EN := "SR Blackword Step motor No.3 เบิกจ่าย 15",
                  Output => "Output ปุ่มยืนยันหน้า Screen",
                  ENO => #_w44);
   #_w46 := #_w44 AND "Output ปุ่มยืนยันหน้า Screen";
   "ตัวเลือกยา (20)"("ปึ่ม 1" := "ยา 16",
                     "ปึ่ม 2" := "ยา 42",
                     "ปึ่ม 3" := "ยา 68",
                     "ปึ่ม 4" := "ยา 94",
                     "ปึ่ม 5" := "ยา 120",
                     "ปึ่ม 6" := "ยา 146",
                     "ปึ่ม 7" := "ยา 172",
                     "ปึ่ม 8" := "ยา 198",
                     "ปึ่ม 9" := "ยา 224",
                     "ปึ่ม 10" := "ยา 250",
                     "ปึ่ม 11" := "ยา 276",
                     "ปึ่ม 12" := "ยา 302",
                     "ปึ่ม 13" := "ยา 328",
                     "ปึ่ม 14" := "ยา 354",
                     "ปึ่ม 15" := "ยา 380",
                     "ปึ่ม 16" := "ยา 406",
                     "ปึ่ม 17" := "ยา 432",
                     "ปึ่ม 18" := "ยา 458",
                     "ปึ่ม 19" := "ยา 484",
                     "ปึ่ม 20" := "ยา 510",
                     "เมื่อกดปุ่ม" => "Output Blackword Step motor No.3 เบิกจ่าย 16",
                     ENO => #_w45);
   IF #_w45 AND "Output Blackword Step motor No.3 เบิกจ่าย 16" THEN
       "SR Blackword Step motor No.3 เบิกจ่าย 16" := TRUE;   // SR flip-flop
   END_IF;
   IF "Output black No3 16" OR "ปุ่มClear" THEN "SR Blackword Step motor No.3 เบิกจ่าย 16" := FALSE; END_IF;
   "button start"(EN := "SR Blackword Step motor No.3 เบิกจ่าย 16",
                  Output => "Output ปุ่มยืนยันหน้า Screen",
                  ENO => #_w47);
   #_w49 := #_w47 AND "Output ปุ่มยืนยันหน้า Screen";
   "ตัวเลือกยา (20)"("ปึ่ม 1" := "ยา 17",
                     "ปึ่ม 2" := "ยา 43",
                     "ปึ่ม 3" := "ยา 69",
                     "ปึ่ม 4" := "ยา 95",
                     "ปึ่ม 5" := "ยา 121",
                     "ปึ่ม 6" := "ยา 147",
                     "ปึ่ม 7" := "ยา 173",
                     "ปึ่ม 8" := "ยา 199",
                     "ปึ่ม 9" := "ยา 225",
                     "ปึ่ม 10" := "ยา 251",
                     "ปึ่ม 11" := "ยา 277",
                     "ปึ่ม 12" := "ยา 303",
                     "ปึ่ม 13" := "ยา 329",
                     "ปึ่ม 14" := "ยา 355",
                     "ปึ่ม 15" := "ยา 381",
                     "ปึ่ม 16" := "ยา 407",
                     "ปึ่ม 17" := "ยา 433",
                     "ปึ่ม 18" := "ยา 459",
                     "ปึ่ม 19" := "ยา 485",
                     "ปึ่ม 20" := "ยา 511",
                     "เมื่อกดปุ่ม" => "Output Blackword Step motor No.3 เบิกจ่าย 17",
                     ENO => #_w48);
   IF #_w48 AND "Output Blackword Step motor No.3 เบิกจ่าย 17" THEN
       "SR Blackword Step motor No.3 เบิกจ่าย 17" := TRUE;   // SR flip-flop
   END_IF;
   IF "Output black No3 17" OR "ปุ่มClear" THEN "SR Blackword Step motor No.3 เบิกจ่าย 17" := FALSE; END_IF;
   "button start"(EN := "SR Blackword Step motor No.3 เบิกจ่าย 17",
                  Output => "Output ปุ่มยืนยันหน้า Screen",
                  ENO => #_w50);
   #_w52 := #_w50 AND "Output ปุ่มยืนยันหน้า Screen";
   "ตัวเลือกยา (20)"("ปึ่ม 1" := "ยา 18",
                     "ปึ่ม 2" := "ยา 44",
                     "ปึ่ม 3" := "ยา 70",
                     "ปึ่ม 4" := "ยา 96",
                     "ปึ่ม 5" := "ยา 122",
                     "ปึ่ม 6" := "ยา 148",
                     "ปึ่ม 7" := "ยา 174",
                     "ปึ่ม 8" := "ยา 200",
                     "ปึ่ม 9" := "ยา 226",
                     "ปึ่ม 10" := "ยา 252",
                     "ปึ่ม 11" := "ยา 278",
                     "ปึ่ม 12" := "ยา 304",
                     "ปึ่ม 13" := "ยา 330",
                     "ปึ่ม 14" := "ยา 356",
                     "ปึ่ม 15" := "ยา 382",
                     "ปึ่ม 16" := "ยา 408",
                     "ปึ่ม 17" := "ยา 434",
                     "ปึ่ม 18" := "ยา 460",
                     "ปึ่ม 19" := "ยา 486",
                     "ปึ่ม 20" := "ยา 512",
                     "เมื่อกดปุ่ม" => "Output Blackword Step motor No.3 เบิกจ่าย 18",
                     ENO => #_w51);
   IF #_w51 AND "Output Blackword Step motor No.3 เบิกจ่าย 18" THEN
       "SR Blackword Step motor No.3 เบิกจ่าย 18" := TRUE;   // SR flip-flop
   END_IF;
   IF "Output black No3 18" OR "ปุ่มClear" THEN "SR Blackword Step motor No.3 เบิกจ่าย 18" := FALSE; END_IF;
   "button start"(EN := "SR Blackword Step motor No.3 เบิกจ่าย 18",
                  Output => "Output ปุ่มยืนยันหน้า Screen",
                  ENO => #_w53);
   #_w55 := #_w53 AND "Output ปุ่มยืนยันหน้า Screen";
   "ตัวเลือกยา (20)"("ปึ่ม 1" := "ยา 19",
                     "ปึ่ม 2" := "ยา 45",
                     "ปึ่ม 3" := "ยา 71",
                     "ปึ่ม 4" := "ยา 97",
                     "ปึ่ม 5" := "ยา 123",
                     "ปึ่ม 6" := "ยา 149",
                     "ปึ่ม 7" := "ยา 175",
                     "ปึ่ม 8" := "ยา 201",
                     "ปึ่ม 9" := "ยา 227",
                     "ปึ่ม 10" := "ยา 253",
                     "ปึ่ม 11" := "ยา 279",
                     "ปึ่ม 12" := "ยา 305",
                     "ปึ่ม 13" := "ยา 331",
                     "ปึ่ม 14" := "ยา 357",
                     "ปึ่ม 15" := "ยา 383",
                     "ปึ่ม 16" := "ยา 409",
                     "ปึ่ม 17" := "ยา 435",
                     "ปึ่ม 18" := "ยา 461",
                     "ปึ่ม 19" := "ยา 487",
                     "ปึ่ม 20" := "ยา 513",
                     "เมื่อกดปุ่ม" => "Output Blackword Step motor No.3 เบิกจ่าย 19",
                     ENO => #_w54);
   IF #_w54 AND "Output Blackword Step motor No.3 เบิกจ่าย 19" THEN
       "SR Blackword Step motor No.3 เบิกจ่าย 19" := TRUE;   // SR flip-flop
   END_IF;
   IF "Output black No3 19" OR "ปุ่มClear" THEN "SR Blackword Step motor No.3 เบิกจ่าย 19" := FALSE; END_IF;
   "button start"(EN := "SR Blackword Step motor No.3 เบิกจ่าย 19",
                  Output => "Output ปุ่มยืนยันหน้า Screen",
                  ENO => #_w56);
   #_w58 := #_w56 AND "Output ปุ่มยืนยันหน้า Screen";
   "ตัวเลือกยา (20)"("ปึ่ม 1" := "ยา 20",
                     "ปึ่ม 2" := "ยา 46",
                     "ปึ่ม 3" := "ยา 72",
                     "ปึ่ม 4" := "ยา 98",
                     "ปึ่ม 5" := "ยา 124",
                     "ปึ่ม 6" := "ยา 150",
                     "ปึ่ม 7" := "ยา 176",
                     "ปึ่ม 8" := "ยา 202",
                     "ปึ่ม 9" := "ยา 228",
                     "ปึ่ม 10" := "ยา 254",
                     "ปึ่ม 11" := "ยา 280",
                     "ปึ่ม 12" := "ยา 306",
                     "ปึ่ม 13" := "ยา 332",
                     "ปึ่ม 14" := "ยา 358",
                     "ปึ่ม 15" := "ยา 384",
                     "ปึ่ม 16" := "ยา 410",
                     "ปึ่ม 17" := "ยา 436",
                     "ปึ่ม 18" := "ยา 462",
                     "ปึ่ม 19" := "ยา 488",
                     "ปึ่ม 20" := "ยา 514",
                     "เมื่อกดปุ่ม" => "Output Blackword Step motor No.3 เบิกจ่าย 20",
                     ENO => #_w57);
   IF #_w57 AND "Output Blackword Step motor No.3 เบิกจ่าย 20" THEN
       "SR Blackword Step motor No.3 เบิกจ่าย 20" := TRUE;   // SR flip-flop
   END_IF;
   IF "Output black No3 20" OR "ปุ่มClear" THEN "SR Blackword Step motor No.3 เบิกจ่าย 20" := FALSE; END_IF;
   "button start"(EN := "SR Blackword Step motor No.3 เบิกจ่าย 20",
                  Output => "Output ปุ่มยืนยันหน้า Screen",
                  ENO => #_w59);
   #_w61 := #_w59 AND "Output ปุ่มยืนยันหน้า Screen";
   "ตัวเลือกยา (20)"("ปึ่ม 1" := "ยา 21",
                     "ปึ่ม 2" := "ยา 47",
                     "ปึ่ม 3" := "ยา 73",
                     "ปึ่ม 4" := "ยา 99",
                     "ปึ่ม 5" := "ยา 125",
                     "ปึ่ม 6" := "ยา 151",
                     "ปึ่ม 7" := "ยา 177",
                     "ปึ่ม 8" := "ยา 203",
                     "ปึ่ม 9" := "ยา 229",
                     "ปึ่ม 10" := "ยา 255",
                     "ปึ่ม 11" := "ยา 281",
                     "ปึ่ม 12" := "ยา 307",
                     "ปึ่ม 13" := "ยา 333",
                     "ปึ่ม 14" := "ยา 359",
                     "ปึ่ม 15" := "ยา 385",
                     "ปึ่ม 16" := "ยา 411",
                     "ปึ่ม 17" := "ยา 437",
                     "ปึ่ม 18" := "ยา 463",
                     "ปึ่ม 19" := "ยา 489",
                     "ปึ่ม 20" := "ยา 515",
                     "เมื่อกดปุ่ม" => "Output Blackword Step motor No.3 เบิกจ่าย 21",
                     ENO => #_w60);
   IF #_w60 AND "Output Blackword Step motor No.3 เบิกจ่าย 21" THEN
       "SR Blackword Step motor No.3 เบิกจ่าย 21" := TRUE;   // SR flip-flop
   END_IF;
   IF "Output black No3 21" OR "ปุ่มClear" THEN "SR Blackword Step motor No.3 เบิกจ่าย 21" := FALSE; END_IF;
   "button start"(EN := "SR Blackword Step motor No.3 เบิกจ่าย 21",
                  Output => "Output ปุ่มยืนยันหน้า Screen",
                  ENO => #_w62);
   #_w64 := #_w62 AND "Output ปุ่มยืนยันหน้า Screen";
   "ตัวเลือกยา (20)"("ปึ่ม 1" := "ยา 22",
                     "ปึ่ม 2" := "ยา 48",
                     "ปึ่ม 3" := "ยา 74",
                     "ปึ่ม 4" := "ยา 100",
                     "ปึ่ม 5" := "ยา 126",
                     "ปึ่ม 6" := "ยา 152",
                     "ปึ่ม 7" := "ยา 178",
                     "ปึ่ม 8" := "ยา 204",
                     "ปึ่ม 9" := "ยา 230",
                     "ปึ่ม 10" := "ยา 256",
                     "ปึ่ม 11" := "ยา 282",
                     "ปึ่ม 12" := "ยา 308",
                     "ปึ่ม 13" := "ยา 334",
                     "ปึ่ม 14" := "ยา 360",
                     "ปึ่ม 15" := "ยา 386",
                     "ปึ่ม 16" := "ยา 412",
                     "ปึ่ม 17" := "ยา 438",
                     "ปึ่ม 18" := "ยา 464",
                     "ปึ่ม 19" := "ยา 490",
                     "ปึ่ม 20" := "ยา 512",
                     "เมื่อกดปุ่ม" => "Output Blackword Step motor No.3 เบิกจ่าย 22",
                     ENO => #_w63);
   IF #_w63 AND "Output Blackword Step motor No.3 เบิกจ่าย 22" THEN
       "SR Blackword Step motor No.3 เบิกจ่าย 22" := TRUE;   // SR flip-flop
   END_IF;
   IF "Output black No3 22" OR "ปุ่มClear" THEN "SR Blackword Step motor No.3 เบิกจ่าย 22" := FALSE; END_IF;
   "button start"(EN := "SR Blackword Step motor No.3 เบิกจ่าย 22",
                  Output => "Output ปุ่มยืนยันหน้า Screen",
                  ENO => #_w65);
   #_w67 := #_w65 AND "Output ปุ่มยืนยันหน้า Screen";
   "ตัวเลือกยา (20)"("ปึ่ม 1" := "ยา 23",
                     "ปึ่ม 2" := "ยา 49",
                     "ปึ่ม 3" := "ยา 75",
                     "ปึ่ม 4" := "ยา 101",
                     "ปึ่ม 5" := "ยา 127",
                     "ปึ่ม 6" := "ยา 153",
                     "ปึ่ม 7" := "ยา 179",
                     "ปึ่ม 8" := "ยา 205",
                     "ปึ่ม 9" := "ยา 231",
                     "ปึ่ม 10" := "ยา 257",
                     "ปึ่ม 11" := "ยา 283",
                     "ปึ่ม 12" := "ยา 309",
                     "ปึ่ม 13" := "ยา 335",
                     "ปึ่ม 14" := "ยา 361",
                     "ปึ่ม 15" := "ยา 387",
                     "ปึ่ม 16" := "ยา 413",
                     "ปึ่ม 17" := "ยา 439",
                     "ปึ่ม 18" := "ยา 465",
                     "ปึ่ม 19" := "ยา 491",
                     "ปึ่ม 20" := "ยา 517",
                     "เมื่อกดปุ่ม" => "Output Blackword Step motor No.3 เบิกจ่าย 23",
                     ENO => #_w66);
   IF #_w66 AND "Output Blackword Step motor No.3 เบิกจ่าย 23" THEN
       "SR Blackword Step motor No.3 เบิกจ่าย 23" := TRUE;   // SR flip-flop
   END_IF;
   IF "Output black No3 23" OR "ปุ่มClear" THEN "SR Blackword Step motor No.3 เบิกจ่าย 23" := FALSE; END_IF;
   "button start"(EN := "SR Blackword Step motor No.3 เบิกจ่าย 23",
                  Output => "Output ปุ่มยืนยันหน้า Screen",
                  ENO => #_w68);
   #_w70 := #_w68 AND "Output ปุ่มยืนยันหน้า Screen";
   "ตัวเลือกยา (20)"("ปึ่ม 1" := "ยา 24",
                     "ปึ่ม 2" := "ยา 50",
                     "ปึ่ม 3" := "ยา 76",
                     "ปึ่ม 4" := "ยา 102",
                     "ปึ่ม 5" := "ยา 128",
                     "ปึ่ม 6" := "ยา 154",
                     "ปึ่ม 7" := "ยา 180",
                     "ปึ่ม 8" := "ยา 206",
                     "ปึ่ม 9" := "ยา 232",
                     "ปึ่ม 10" := "ยา 258",
                     "ปึ่ม 11" := "ยา 284",
                     "ปึ่ม 12" := "ยา 310",
                     "ปึ่ม 13" := "ยา 336",
                     "ปึ่ม 14" := "ยา 362",
                     "ปึ่ม 15" := "ยา 388",
                     "ปึ่ม 16" := "ยา 414",
                     "ปึ่ม 17" := "ยา 440",
                     "ปึ่ม 18" := "ยา 466",
                     "ปึ่ม 19" := "ยา 492",
                     "ปึ่ม 20" := "ยา 518",
                     "เมื่อกดปุ่ม" => "Output Blackword Step motor No.3 เบิกจ่าย 24",
                     ENO => #_w69);
   IF #_w69 AND "Output Blackword Step motor No.3 เบิกจ่าย 24" THEN
       "SR Blackword Step motor No.3 เบิกจ่าย 24" := TRUE;   // SR flip-flop
   END_IF;
   IF "Output black No3 24" OR "ปุ่มClear" THEN "SR Blackword Step motor No.3 เบิกจ่าย 24" := FALSE; END_IF;
   "button start"(EN := "SR Blackword Step motor No.3 เบิกจ่าย 24",
                  Output => "Output ปุ่มยืนยันหน้า Screen",
                  ENO => #_w71);
   #_w73 := #_w71 AND "Output ปุ่มยืนยันหน้า Screen";
   "ตัวเลือกยา (20)"("ปึ่ม 1" := "ยา 25",
                     "ปึ่ม 2" := "ยา 51",
                     "ปึ่ม 3" := "ยา 77",
                     "ปึ่ม 4" := "ยา 103",
                     "ปึ่ม 5" := "ยา 129",
                     "ปึ่ม 6" := "ยา 155",
                     "ปึ่ม 7" := "ยา 181",
                     "ปึ่ม 8" := "ยา 207",
                     "ปึ่ม 9" := "ยา 233",
                     "ปึ่ม 10" := "ยา 259",
                     "ปึ่ม 11" := "ยา 285",
                     "ปึ่ม 12" := "ยา 311",
                     "ปึ่ม 13" := "ยา 337",
                     "ปึ่ม 14" := "ยา 363",
                     "ปึ่ม 15" := "ยา 389",
                     "ปึ่ม 16" := "ยา 415",
                     "ปึ่ม 17" := "ยา 441",
                     "ปึ่ม 18" := "ยา 467",
                     "ปึ่ม 19" := "ยา 493",
                     "ปึ่ม 20" := "ยา 519",
                     "เมื่อกดปุ่ม" => "Output Blackword Step motor No.3 เบิกจ่าย 25",
                     ENO => #_w72);
   IF #_w72 AND "Output Blackword Step motor No.3 เบิกจ่าย 25" THEN
       "SR Blackword Step motor No.3 เบิกจ่าย 25" := TRUE;   // SR flip-flop
   END_IF;
   IF "Output black No3 25" OR "ปุ่มClear" THEN "SR Blackword Step motor No.3 เบิกจ่าย 25" := FALSE; END_IF;
   "button start"(EN := "SR Blackword Step motor No.3 เบิกจ่าย 25",
                  Output => "Output ปุ่มยืนยันหน้า Screen",
                  ENO => #_w74);
   #_w76 := #_w74 AND "Output ปุ่มยืนยันหน้า Screen";
   "ตัวเลือกยา (20)"("ปึ่ม 1" := "ยา 26",
                     "ปึ่ม 2" := "ยา 52",
                     "ปึ่ม 3" := "ยา 78",
                     "ปึ่ม 4" := "ยา 104",
                     "ปึ่ม 5" := "ยา 130",
                     "ปึ่ม 6" := "ยา 156",
                     "ปึ่ม 7" := "ยา 182",
                     "ปึ่ม 8" := "ยา 208",
                     "ปึ่ม 9" := "ยา 234",
                     "ปึ่ม 10" := "ยา 260",
                     "ปึ่ม 11" := "ยา 286",
                     "ปึ่ม 12" := "ยา 312",
                     "ปึ่ม 13" := "ยา 338",
                     "ปึ่ม 14" := "ยา 364",
                     "ปึ่ม 15" := "ยา 390",
                     "ปึ่ม 16" := "ยา 416",
                     "ปึ่ม 17" := "ยา 442",
                     "ปึ่ม 18" := "ยา 468",
                     "ปึ่ม 19" := "ยา 494",
                     "ปึ่ม 20" := "ยา 520",
                     "เมื่อกดปุ่ม" => "Output Blackword Step motor No.3 เบิกจ่าย 26",
                     ENO => #_w75);
   IF #_w75 AND "Output Blackword Step motor No.3 เบิกจ่าย 26" THEN
       "SR Blackword Step motor No.3 เบิกจ่าย 26" := TRUE;   // SR flip-flop
   END_IF;
   IF "Output black No3 26" OR "ปุ่มClear" THEN "SR Blackword Step motor No.3 เบิกจ่าย 26" := FALSE; END_IF;
   "button start"(EN := "SR Blackword Step motor No.3 เบิกจ่าย 26",
                  Output => "Output ปุ่มยืนยันหน้า Screen",
                  ENO => #_w77);
   "IEC_Counter_0_DB_1597".CTU(CU := (#_w4 OR #_w7 OR #_w10 OR #_w13 OR #_w16 OR #_w19 OR #_w22 OR #_w25 OR #_w28 OR #_w31 OR #_w34 OR #_w37 OR #_w40 OR #_w43 OR #_w46 OR #_w49 OR #_w52 OR #_w55 OR #_w58 OR #_w61 OR #_w64 OR #_w67 OR #_w70 OR #_w73 OR #_w76 OR (#_w77 AND "Output ปุ่มยืนยันหน้า Screen")) AND (("SR Step Motro 3  เบิกจ่าย 1" AND ("IEC_Timer_0_DB_100".ET = T#1.75s)) OR ("SR Step Motro 3  เบิกจ่าย 2" AND ("IEC_Timer_0_DB_101".ET = T#1.2s)) OR ("SR Step Motro 3  เบิกจ่าย 3" AND ("IEC_Timer_0_DB_102".ET = T#1s)) OR ("SR Step Motro 3  เบิกจ่าย 4" AND ("IEC_Timer_0_DB_103".ET = T#0.8s)) OR ("SR Step Motro 3  เบิกจ่าย 5" AND ("IEC_Timer_0_DB_104".ET = T#0.6s)) OR ("SR Step Motro 3  เบิกจ่าย 6" AND ("IEC_Timer_0_DB_105".ET = T#0.4s)) OR ("SR Step Motro 3  เบิกจ่าย 7" AND ("IEC_Timer_0_DB_106".ET = T#0.2s)) OR ("SR Step Motro 3  เบิกจ่าย 8" AND ("IEC_Timer_0_DB_107".ET = T#0.2s)) OR ("SR Step Motro 3  เบิกจ่าย 9" AND ("IEC_Timer_0_DB_108".ET = T#0.2s)) OR ("SR Step Motro 3  เบิกจ่าย 10" AND ("IEC_Timer_0_DB_109".ET = T#0.4s)) OR ("SR Step Motro 3  เบิกจ่าย 11" AND ("IEC_Timer_0_DB_110".ET = T#0.6s)) OR ("SR Step Motro 3  เบิกจ่าย 12" AND ("IEC_Timer_0_DB_111".ET = T#0.8s)) OR ("SR Step Motro 3  เบิกจ่าย 13" AND ("IEC_Timer_0_DB_112".ET = T#1s)) OR ("SR Step Motro 3  เบิกจ่าย 14" AND ("IEC_Timer_0_DB_113".ET = T#1.2s)) OR ("SR Step Motro 3  เบิกจ่าย 15" AND ("IEC_Timer_0_DB_114".ET = T#1.4s)) OR ("SR Step Motro 3  เบิกจ่าย 16" AND ("IEC_Timer_0_DB_115".ET = T#1.6s)) OR ("SR Step Motro 3  เบิกจ่าย 17" AND ("IEC_Timer_0_DB_116".ET = T#1.8s)) OR ("SR Step Motro 3  เบิกจ่าย 18" AND ("IEC_Timer_0_DB_117".ET = T#2s)) OR ("SR Step Motro 3  เบิกจ่าย 19" AND ("IEC_Timer_0_DB_118".ET = T#2.2s)) OR ("SR Step Motro 3  เบิกจ่าย 20" AND ("IEC_Timer_0_DB_119".ET = T#2.4s))),
                           R := "เวลาหลังจากเคลื่อนที่ถึงตำแหน่งเป้าหมาย (26) Blackword",
                           PV := 1);
   #"Stepper Motor  ทำงาน3" := "IEC_Counter_0_DB_1597".Q;
END_REGION

REGION Network 2
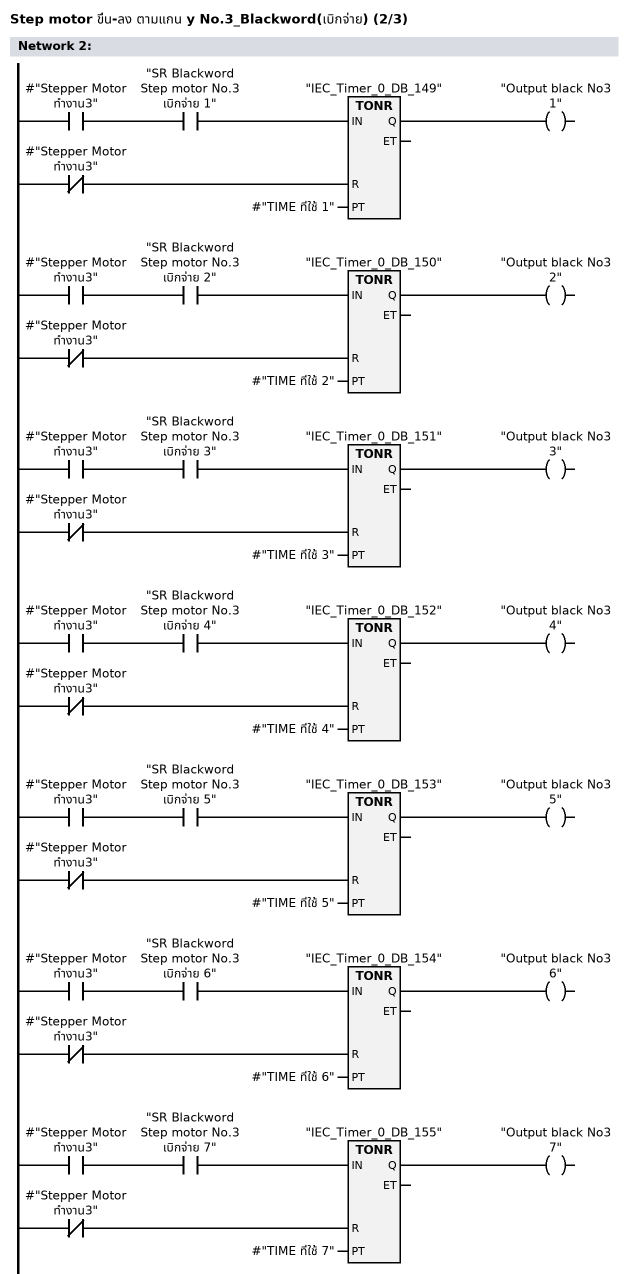
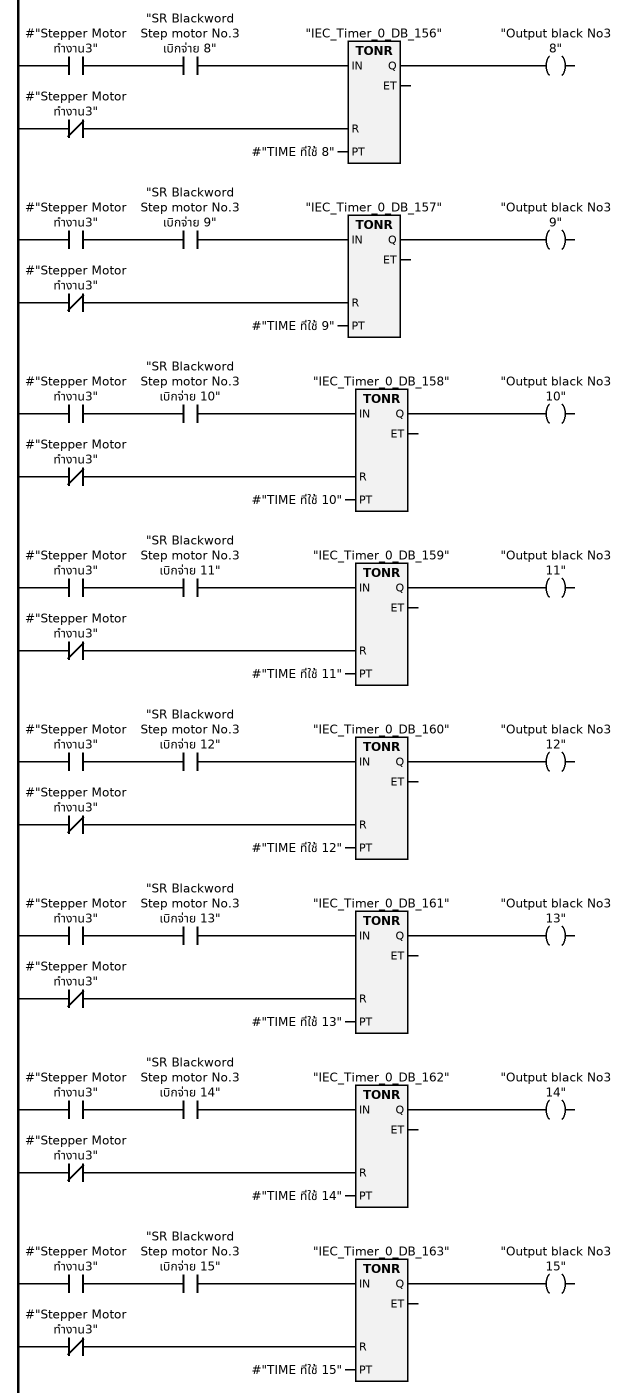
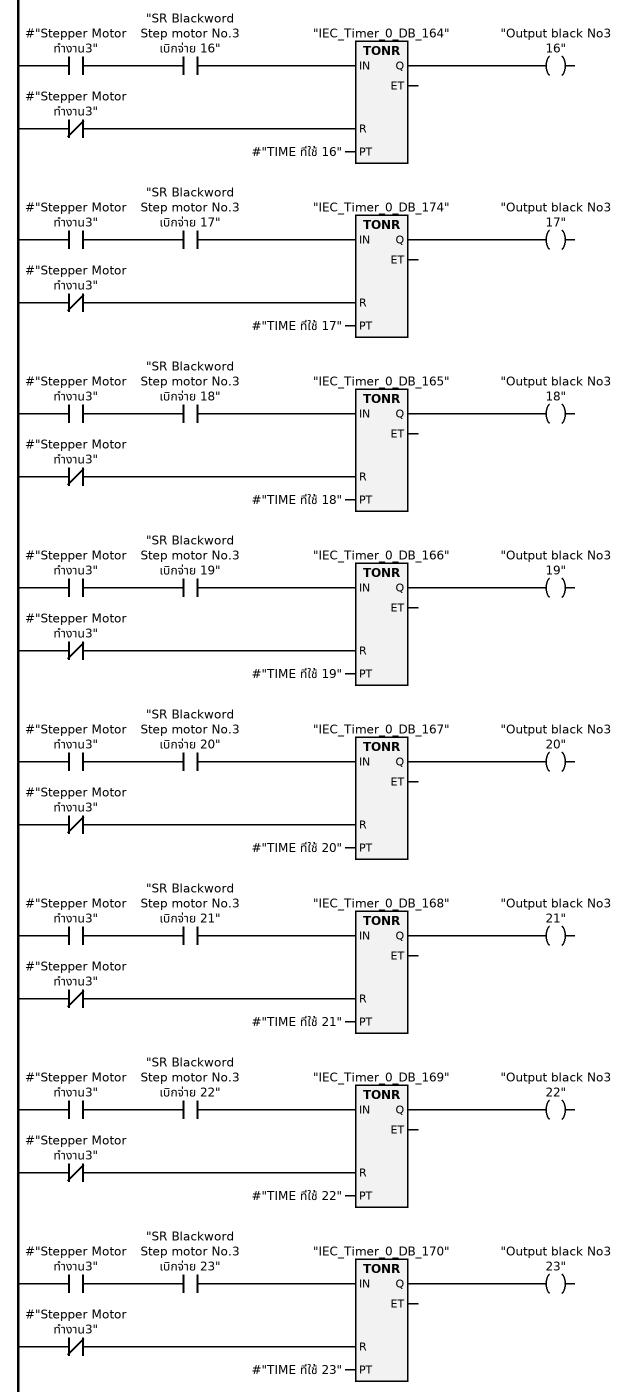
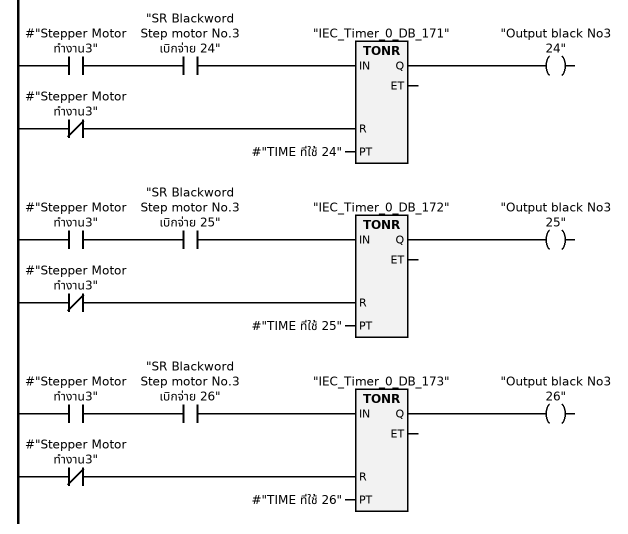
   "IEC_Timer_0_DB_149".TONR(IN := #"Stepper Motor  ทำงาน3" AND "SR Blackword Step motor No.3 เบิกจ่าย 1",
                           R := NOT #"Stepper Motor  ทำงาน3",
                           PT := #"TIME ที่ใช้ 1");
   "Output black No3 1" := "IEC_Timer_0_DB_149".Q;
   "IEC_Timer_0_DB_150".TONR(IN := #"Stepper Motor  ทำงาน3" AND "SR Blackword Step motor No.3 เบิกจ่าย 2",
                           R := NOT #"Stepper Motor  ทำงาน3",
                           PT := #"TIME ที่ใช้ 2");
   "Output black No3 2" := "IEC_Timer_0_DB_150".Q;
   "IEC_Timer_0_DB_151".TONR(IN := #"Stepper Motor  ทำงาน3" AND "SR Blackword Step motor No.3 เบิกจ่าย 3",
                           R := NOT #"Stepper Motor  ทำงาน3",
                           PT := #"TIME ที่ใช้ 3");
   "Output black No3 3" := "IEC_Timer_0_DB_151".Q;
   "IEC_Timer_0_DB_152".TONR(IN := #"Stepper Motor  ทำงาน3" AND "SR Blackword Step motor No.3 เบิกจ่าย 4",
                           R := NOT #"Stepper Motor  ทำงาน3",
                           PT := #"TIME ที่ใช้ 4");
   "Output black No3 4" := "IEC_Timer_0_DB_152".Q;
   "IEC_Timer_0_DB_153".TONR(IN := #"Stepper Motor  ทำงาน3" AND "SR Blackword Step motor No.3 เบิกจ่าย 5",
                           R := NOT #"Stepper Motor  ทำงาน3",
                           PT := #"TIME ที่ใช้ 5");
   "Output black No3 5" := "IEC_Timer_0_DB_153".Q;
   "IEC_Timer_0_DB_154".TONR(IN := #"Stepper Motor  ทำงาน3" AND "SR Blackword Step motor No.3 เบิกจ่าย 6",
                           R := NOT #"Stepper Motor  ทำงาน3",
                           PT := #"TIME ที่ใช้ 6");
   "Output black No3 6" := "IEC_Timer_0_DB_154".Q;
   "IEC_Timer_0_DB_155".TONR(IN := #"Stepper Motor  ทำงาน3" AND "SR Blackword Step motor No.3 เบิกจ่าย 7",
                           R := NOT #"Stepper Motor  ทำงาน3",
                           PT := #"TIME ที่ใช้ 7");
   "Output black No3 7" := "IEC_Timer_0_DB_155".Q;
   "IEC_Timer_0_DB_156".TONR(IN := #"Stepper Motor  ทำงาน3" AND "SR Blackword Step motor No.3 เบิกจ่าย 8",
                           R := NOT #"Stepper Motor  ทำงาน3",
                           PT := #"TIME ที่ใช้ 8");
   "Output black No3 8" := "IEC_Timer_0_DB_156".Q;
   "IEC_Timer_0_DB_157".TONR(IN := #"Stepper Motor  ทำงาน3" AND "SR Blackword Step motor No.3 เบิกจ่าย 9",
                           R := NOT #"Stepper Motor  ทำงาน3",
                           PT := #"TIME ที่ใช้ 9");
   "Output black No3 9" := "IEC_Timer_0_DB_157".Q;
   "IEC_Timer_0_DB_158".TONR(IN := #"Stepper Motor  ทำงาน3" AND "SR Blackword Step motor No.3 เบิกจ่าย 10",
                           R := NOT #"Stepper Motor  ทำงาน3",
                           PT := #"TIME ที่ใช้ 10");
   "Output black No3 10" := "IEC_Timer_0_DB_158".Q;
   "IEC_Timer_0_DB_159".TONR(IN := #"Stepper Motor  ทำงาน3" AND "SR Blackword Step motor No.3 เบิกจ่าย 11",
                           R := NOT #"Stepper Motor  ทำงาน3",
                           PT := #"TIME ที่ใช้ 11");
   "Output black No3 11" := "IEC_Timer_0_DB_159".Q;
   "IEC_Timer_0_DB_160".TONR(IN := #"Stepper Motor  ทำงาน3" AND "SR Blackword Step motor No.3 เบิกจ่าย 12",
                           R := NOT #"Stepper Motor  ทำงาน3",
                           PT := #"TIME ที่ใช้ 12");
   "Output black No3 12" := "IEC_Timer_0_DB_160".Q;
   "IEC_Timer_0_DB_161".TONR(IN := #"Stepper Motor  ทำงาน3" AND "SR Blackword Step motor No.3 เบิกจ่าย 13",
                           R := NOT #"Stepper Motor  ทำงาน3",
                           PT := #"TIME ที่ใช้ 13");
   "Output black No3 13" := "IEC_Timer_0_DB_161".Q;
   "IEC_Timer_0_DB_162".TONR(IN := #"Stepper Motor  ทำงาน3" AND "SR Blackword Step motor No.3 เบิกจ่าย 14",
                           R := NOT #"Stepper Motor  ทำงาน3",
                           PT := #"TIME ที่ใช้ 14");
   "Output black No3 14" := "IEC_Timer_0_DB_162".Q;
   "IEC_Timer_0_DB_163".TONR(IN := #"Stepper Motor  ทำงาน3" AND "SR Blackword Step motor No.3 เบิกจ่าย 15",
                           R := NOT #"Stepper Motor  ทำงาน3",
                           PT := #"TIME ที่ใช้ 15");
   "Output black No3 15" := "IEC_Timer_0_DB_163".Q;
   "IEC_Timer_0_DB_164".TONR(IN := #"Stepper Motor  ทำงาน3" AND "SR Blackword Step motor No.3 เบิกจ่าย 16",
                           R := NOT #"Stepper Motor  ทำงาน3",
                           PT := #"TIME ที่ใช้ 16");
   "Output black No3 16" := "IEC_Timer_0_DB_164".Q;
   "IEC_Timer_0_DB_174".TONR(IN := #"Stepper Motor  ทำงาน3" AND "SR Blackword Step motor No.3 เบิกจ่าย 17",
                           R := NOT #"Stepper Motor  ทำงาน3",
                           PT := #"TIME ที่ใช้ 17");
   "Output black No3 17" := "IEC_Timer_0_DB_174".Q;
   "IEC_Timer_0_DB_165".TONR(IN := #"Stepper Motor  ทำงาน3" AND "SR Blackword Step motor No.3 เบิกจ่าย 18",
                           R := NOT #"Stepper Motor  ทำงาน3",
                           PT := #"TIME ที่ใช้ 18");
   "Output black No3 18" := "IEC_Timer_0_DB_165".Q;
   "IEC_Timer_0_DB_166".TONR(IN := #"Stepper Motor  ทำงาน3" AND "SR Blackword Step motor No.3 เบิกจ่าย 19",
                           R := NOT #"Stepper Motor  ทำงาน3",
                           PT := #"TIME ที่ใช้ 19");
   "Output black No3 19" := "IEC_Timer_0_DB_166".Q;
   "IEC_Timer_0_DB_167".TONR(IN := #"Stepper Motor  ทำงาน3" AND "SR Blackword Step motor No.3 เบิกจ่าย 20",
                           R := NOT #"Stepper Motor  ทำงาน3",
                           PT := #"TIME ที่ใช้ 20");
   "Output black No3 20" := "IEC_Timer_0_DB_167".Q;
   "IEC_Timer_0_DB_168".TONR(IN := #"Stepper Motor  ทำงาน3" AND "SR Blackword Step motor No.3 เบิกจ่าย 21",
                           R := NOT #"Stepper Motor  ทำงาน3",
                           PT := #"TIME ที่ใช้ 21");
   "Output black No3 21" := "IEC_Timer_0_DB_168".Q;
   "IEC_Timer_0_DB_169".TONR(IN := #"Stepper Motor  ทำงาน3" AND "SR Blackword Step motor No.3 เบิกจ่าย 22",
                           R := NOT #"Stepper Motor  ทำงาน3",
                           PT := #"TIME ที่ใช้ 22");
   "Output black No3 22" := "IEC_Timer_0_DB_169".Q;
   "IEC_Timer_0_DB_170".TONR(IN := #"Stepper Motor  ทำงาน3" AND "SR Blackword Step motor No.3 เบิกจ่าย 23",
                           R := NOT #"Stepper Motor  ทำงาน3",
                           PT := #"TIME ที่ใช้ 23");
   "Output black No3 23" := "IEC_Timer_0_DB_170".Q;
   "IEC_Timer_0_DB_171".TONR(IN := #"Stepper Motor  ทำงาน3" AND "SR Blackword Step motor No.3 เบิกจ่าย 24",
                           R := NOT #"Stepper Motor  ทำงาน3",
                           PT := #"TIME ที่ใช้ 24");
   "Output black No3 24" := "IEC_Timer_0_DB_171".Q;
   "IEC_Timer_0_DB_172".TONR(IN := #"Stepper Motor  ทำงาน3" AND "SR Blackword Step motor No.3 เบิกจ่าย 25",
                           R := NOT #"Stepper Motor  ทำงาน3",
                           PT := #"TIME ที่ใช้ 25");
   "Output black No3 25" := "IEC_Timer_0_DB_172".Q;
   "IEC_Timer_0_DB_173".TONR(IN := #"Stepper Motor  ทำงาน3" AND "SR Blackword Step motor No.3 เบิกจ่าย 26",
                           R := NOT #"Stepper Motor  ทำงาน3",
                           PT := #"TIME ที่ใช้ 26");
   "Output black No3 26" := "IEC_Timer_0_DB_173".Q;
END_REGION

REGION Network 3
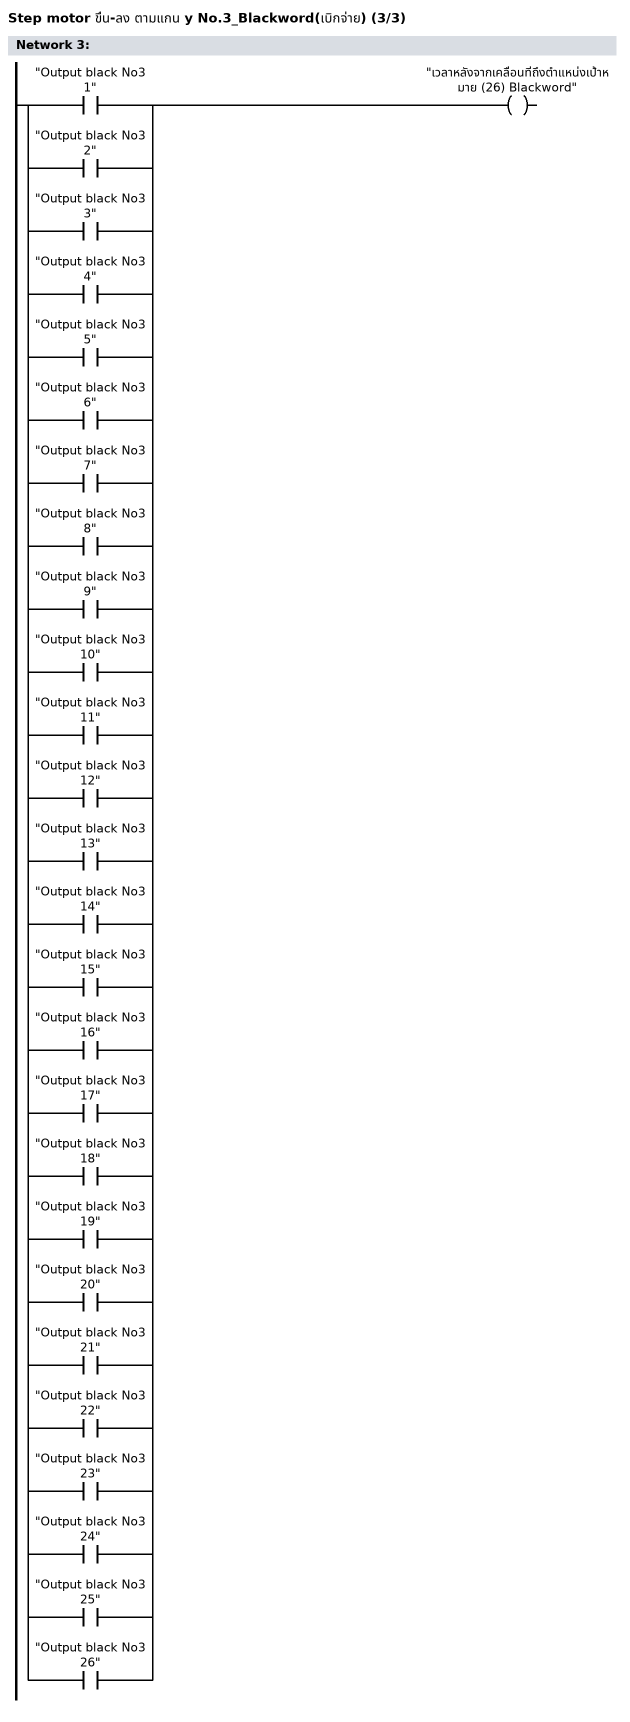
   RUNG wire#powerrail
      Contact( "Output black No3 1" )
      wire#w1
      Coil( "เวลาหลังจากเคลื่อนที่ถึงตำแหน่งเป้าหมาย (26) Blackword" )
   END_RUNG
   RUNG wire#powerrail
      Contact( "Output black No3 2" )
   END_RUNG wire#w1
   RUNG wire#powerrail
      Contact( "Output black No3 3" )
   END_RUNG wire#w1
   RUNG wire#powerrail
      Contact( "Output black No3 4" )
   END_RUNG wire#w1
   RUNG wire#powerrail
      Contact( "Output black No3 5" )
   END_RUNG wire#w1
   RUNG wire#powerrail
      Contact( "Output black No3 6" )
   END_RUNG wire#w1
   RUNG wire#powerrail
      Contact( "Output black No3 7" )
   END_RUNG wire#w1
   RUNG wire#powerrail
      Contact( "Output black No3 8" )
   END_RUNG wire#w1
   RUNG wire#powerrail
      Contact( "Output black No3 9" )
   END_RUNG wire#w1
   RUNG wire#powerrail
      Contact( "Output black No3 10" )
   END_RUNG wire#w1
   RUNG wire#powerrail
      Contact( "Output black No3 11" )
   END_RUNG wire#w1
   RUNG wire#powerrail
      Contact( "Output black No3 12" )
   END_RUNG wire#w1
   RUNG wire#powerrail
      Contact( "Output black No3 13" )
   END_RUNG wire#w1
   RUNG wire#powerrail
      Contact( "Output black No3 14" )
   END_RUNG wire#w1
   RUNG wire#powerrail
      Contact( "Output black No3 15" )
   END_RUNG wire#w1
   RUNG wire#powerrail
      Contact( "Output black No3 16" )
   END_RUNG wire#w1
   RUNG wire#powerrail
      Contact( "Output black No3 17" )
   END_RUNG wire#w1
   RUNG wire#powerrail
      Contact( "Output black No3 18" )
   END_RUNG wire#w1
   RUNG wire#powerrail
      Contact( "Output black No3 19" )
   END_RUNG wire#w1
   RUNG wire#powerrail
      Contact( "Output black No3 20" )
   END_RUNG wire#w1
   RUNG wire#powerrail
      Contact( "Output black No3 21" )
   END_RUNG wire#w1
   RUNG wire#powerrail
      Contact( "Output black No3 22" )
   END_RUNG wire#w1
   RUNG wire#powerrail
      Contact( "Output black No3 23" )
   END_RUNG wire#w1
   RUNG wire#powerrail
      Contact( "Output black No3 24" )
   END_RUNG wire#w1
   RUNG wire#powerrail
      Contact( "Output black No3 25" )
   END_RUNG wire#w1
   RUNG wire#powerrail
      Contact( "Output black No3 26" )
   END_RUNG wire#w1
   // the same network as SCL:
   "เวลาหลังจากเคลื่อนที่ถึงตำแหน่งเป้าหมาย (26) Blackword" := "Output black No3 1" OR "Output black No3 2" OR "Output black No3 3" OR "Output black No3 4" OR "Output black No3 5" OR "Output black No3 6" OR "Output black No3 7" OR "Output black No3 8" OR "Output black No3 9" OR "Output black No3 10" OR "Output black No3 11" OR "Output black No3 12" OR "Output black No3 13" OR "Output black No3 14" OR "Output black No3 15" OR "Output black No3 16" OR "Output black No3 17" OR "Output black No3 18" OR "Output black No3 19" OR "Output black No3 20" OR "Output black No3 21" OR "Output black No3 22" OR "Output black No3 23" OR "Output black No3 24" OR "Output black No3 25" OR "Output black No3 26";
END_REGION
END_FUNCTION_BLOCK

FUNCTION "Test_F" : Void   // FC19, LAD
{ S7_Optimized_Access := 'TRUE' }
VERSION : 0.1
BEGIN

REGION Network 1
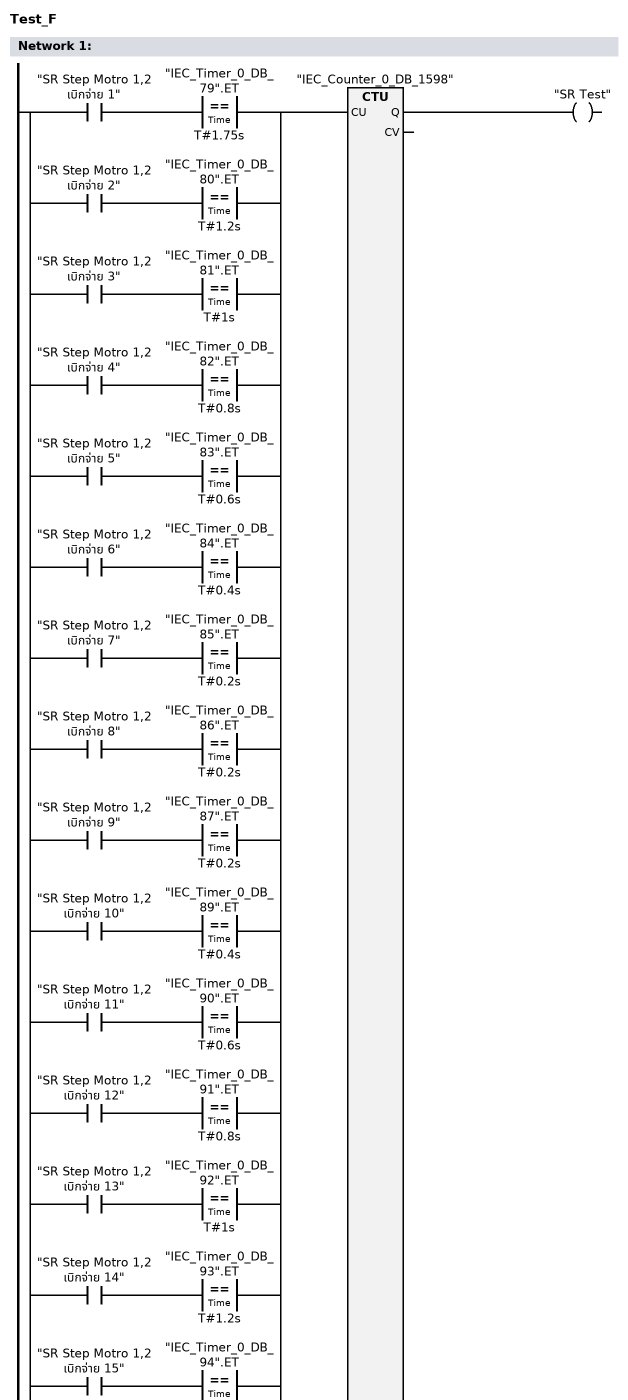
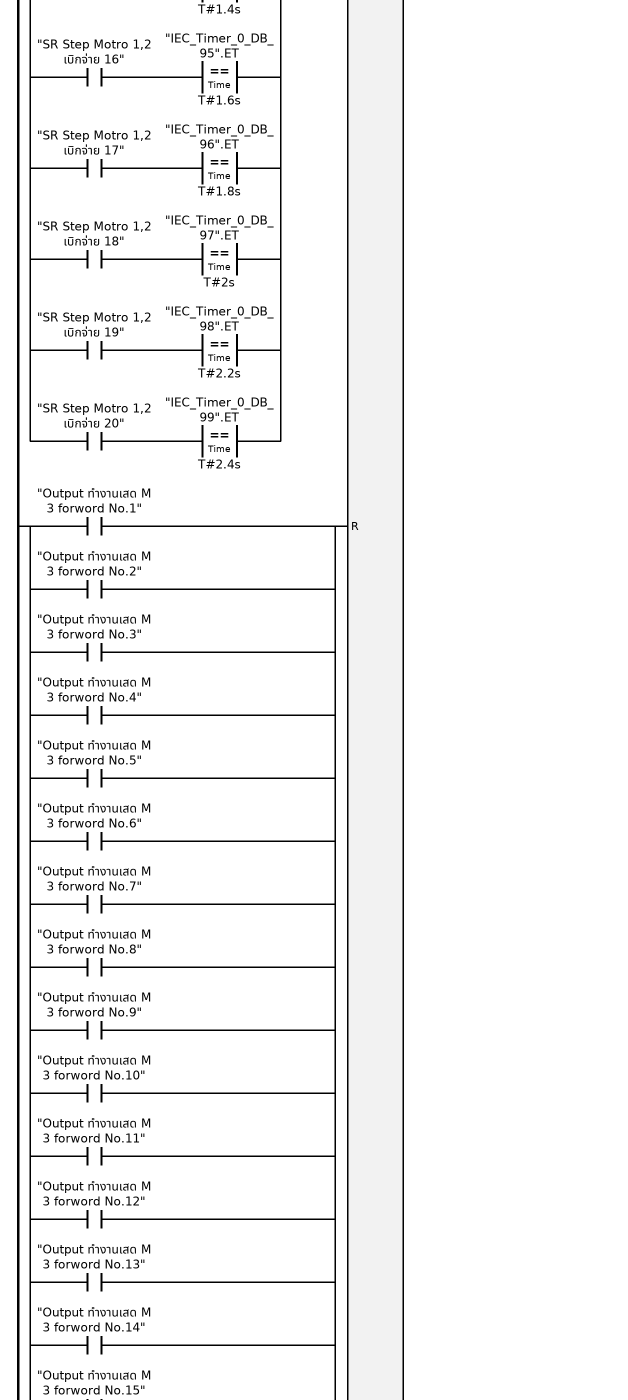
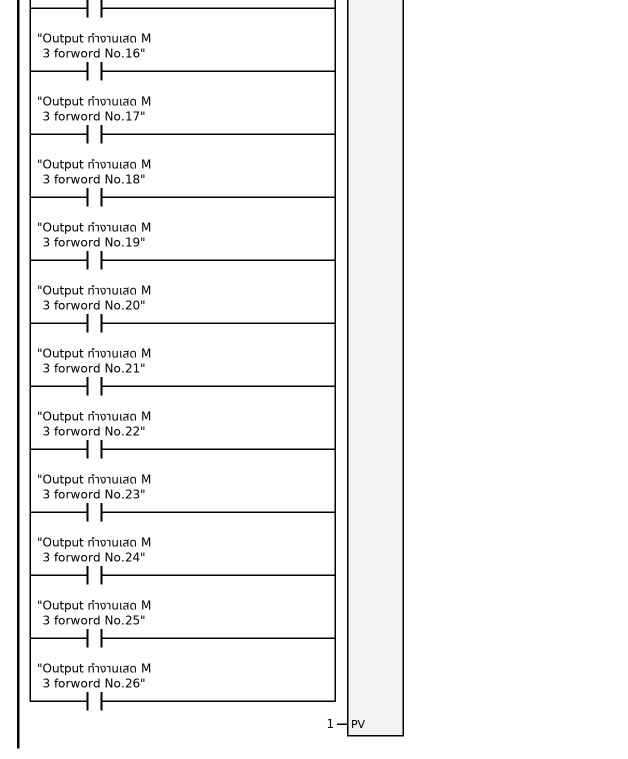
   "IEC_Counter_0_DB_1598".CTU(CU := ("SR Step Motro 1,2  เบิกจ่าย 1" AND ("IEC_Timer_0_DB_79".ET = T#1.75s)) OR ("SR Step Motro 1,2  เบิกจ่าย 2" AND ("IEC_Timer_0_DB_80".ET = T#1.2s)) OR ("SR Step Motro 1,2  เบิกจ่าย 3" AND ("IEC_Timer_0_DB_81".ET = T#1s)) OR ("SR Step Motro 1,2  เบิกจ่าย 4" AND ("IEC_Timer_0_DB_82".ET = T#0.8s)) OR ("SR Step Motro 1,2  เบิกจ่าย 5" AND ("IEC_Timer_0_DB_83".ET = T#0.6s)) OR ("SR Step Motro 1,2  เบิกจ่าย 6" AND ("IEC_Timer_0_DB_84".ET = T#0.4s)) OR ("SR Step Motro 1,2  เบิกจ่าย 7" AND ("IEC_Timer_0_DB_85".ET = T#0.2s)) OR ("SR Step Motro 1,2  เบิกจ่าย 8" AND ("IEC_Timer_0_DB_86".ET = T#0.2s)) OR ("SR Step Motro 1,2  เบิกจ่าย 9" AND ("IEC_Timer_0_DB_87".ET = T#0.2s)) OR ("SR Step Motro 1,2  เบิกจ่าย 10" AND ("IEC_Timer_0_DB_89".ET = T#0.4s)) OR ("SR Step Motro 1,2  เบิกจ่าย 11" AND ("IEC_Timer_0_DB_90".ET = T#0.6s)) OR ("SR Step Motro 1,2  เบิกจ่าย 12" AND ("IEC_Timer_0_DB_91".ET = T#0.8s)) OR ("SR Step Motro 1,2  เบิกจ่าย 13" AND ("IEC_Timer_0_DB_92".ET = T#1s)) OR ("SR Step Motro 1,2  เบิกจ่าย 14" AND ("IEC_Timer_0_DB_93".ET = T#1.2s)) OR ("SR Step Motro 1,2  เบิกจ่าย 15" AND ("IEC_Timer_0_DB_94".ET = T#1.4s)) OR ("SR Step Motro 1,2  เบิกจ่าย 16" AND ("IEC_Timer_0_DB_95".ET = T#1.6s)) OR ("SR Step Motro 1,2  เบิกจ่าย 17" AND ("IEC_Timer_0_DB_96".ET = T#1.8s)) OR ("SR Step Motro 1,2  เบิกจ่าย 18" AND ("IEC_Timer_0_DB_97".ET = T#2s)) OR ("SR Step Motro 1,2  เบิกจ่าย 19" AND ("IEC_Timer_0_DB_98".ET = T#2.2s)) OR ("SR Step Motro 1,2  เบิกจ่าย 20" AND ("IEC_Timer_0_DB_99".ET = T#2.4s)),
                           R := "Output ทำงานเสด M 3 forword No.1" OR "Output ทำงานเสด M 3 forword No.2" OR "Output ทำงานเสด M 3 forword No.3" OR "Output ทำงานเสด M 3 forword No.4" OR "Output ทำงานเสด M 3 forword No.5" OR "Output ทำงานเสด M 3 forword No.6" OR "Output ทำงานเสด M 3 forword No.7" OR "Output ทำงานเสด M 3 forword No.8" OR "Output ทำงานเสด M 3 forword No.9" OR "Output ทำงานเสด M 3 forword No.10" OR "Output ทำงานเสด M 3 forword No.11" OR "Output ทำงานเสด M 3 forword No.12" OR "Output ทำงานเสด M 3 forword No.13" OR "Output ทำงานเสด M 3 forword No.14" OR "Output ทำงานเสด M 3 forword No.15" OR "Output ทำงานเสด M 3 forword No.16" OR "Output ทำงานเสด M 3 forword No.17" OR "Output ทำงานเสด M 3 forword No.18" OR "Output ทำงานเสด M 3 forword No.19" OR "Output ทำงานเสด M 3 forword No.20" OR "Output ทำงานเสด M 3 forword No.21" OR "Output ทำงานเสด M 3 forword No.22" OR "Output ทำงานเสด M 3 forword No.23" OR "Output ทำงานเสด M 3 forword No.24" OR "Output ทำงานเสด M 3 forword No.25" OR "Output ทำงานเสด M 3 forword No.26",
                           PV := 1);
   "SR Test" := "IEC_Counter_0_DB_1598".Q;
END_REGION
END_FUNCTION

(* ===== HMI "HMI_RT_1" =====
system functions are stored by id; their names below are inferred from use
connection "HMI_Connection_1": ETHERNET, S7_1500_OMS

